(* IEC 61131-3 sources: IEC61131-3_ST_SCL_Mutation_Generator/Tests/mutatedCodeTraffic, 85 files *)

(* ---- M097.st ---- *)
FUNCTION_BLOCK TRAFFIC_CTRL

VAR_INPUT
    PedestrianButton1 : BOOL;
    PedestrianButton2 : BOOL;
END_VAR

VAR_OUTPUT
    NorthSouthRed : BOOL;
    NorthSouthYellow : BOOL;
    NorthSouthGreen : BOOL;
    EastWestRed : BOOL;
    EastWestYellow : BOOL;
    EastWestGreen : BOOL;
    PedestrianLight1 : BOOL;
    PedestrianLight2 : BOOL;
END_VAR

VAR
    LightState : INT := 0; (* 0: North-South Green, 1: North-South Yellow, 2: East-West Green, 3: East-West Yellow *)
    PedestrianRequest1 : BOOL := FALSE;
    PedestrianRequest2 : BOOL := FALSE;
    PedestrianCrossing : BOOL := FALSE;
    Timer : TON;
END_VAR

(* Check for pedestrian requests *)
IF PedestrianButton1 THEN
    PedestrianRequest1 := TRUE;
END_IF;

IF PedestrianButton2 THEN
    PedestrianRequest2 := TRUE;
END_IF;

(* Traffic light state machine *)
CASE LightState OF
    0: (* North-South Green *)
        NorthSouthGreen := TRUE;
        EastWestRed := TRUE;
        IF PedestrianRequest1 AND PedestrianRequest2 THEN (* MUTATED: LOGICAL_OP_REPLACE *)
            Timer(IN := TRUE, PT := T#2s); (* Pedestrian crossing grace period *)
            IF Timer.Q THEN
                Timer(IN := FALSE);
                LightState := 1;
            END_IF;
        END_IF;

    1: (* North-South Yellow *)
        NorthSouthYellow := TRUE;
        EastWestRed := TRUE;
        Timer(IN := TRUE, PT := T#2s); (* Yellow light duration *)
        IF Timer.Q THEN
            Timer(IN := FALSE);
            LightState := 2;
        END_IF;

    2: (* East-West Green *)
        EastWestGreen := TRUE;
        NorthSouthRed := TRUE;
        IF PedestrianRequest1 THEN
            PedestrianLight1 := TRUE;
            PedestrianCrossing := TRUE;
        END_IF;
        IF PedestrianRequest2 THEN
            PedestrianLight2 := TRUE;
            PedestrianCrossing := TRUE;
        END_IF;
        IF PedestrianCrossing THEN
            Timer(IN := TRUE, PT := T#2s); (* Pedestrian crossing period *)
            IF Timer.Q THEN
                Timer(IN := FALSE);
                PedestrianRequest1 := FALSE;
                PedestrianRequest2 := FALSE;
                PedestrianLight1 := FALSE;
                PedestrianLight2 := FALSE;
                PedestrianCrossing := FALSE;
                LightState := 3;
            END_IF;
        END_IF;

    3: (* East-West Yellow *)
        EastWestYellow := TRUE;
        NorthSouthRed := TRUE;
        Timer(IN := TRUE, PT := T#2s); (* Yellow light duration *)
        IF Timer.Q THEN
            Timer(IN := FALSE);
            LightState := 0;
        END_IF;

END_CASE;

END_FUNCTION_BLOCK

(* ---- M098.st ---- *)
FUNCTION_BLOCK TRAFFIC_CTRL

VAR_INPUT
    PedestrianButton1 : BOOL;
    PedestrianButton2 : BOOL;
END_VAR

VAR_OUTPUT
    NorthSouthRed : BOOL;
    NorthSouthYellow : BOOL;
    NorthSouthGreen : BOOL;
    EastWestRed : BOOL;
    EastWestYellow : BOOL;
    EastWestGreen : BOOL;
    PedestrianLight1 : BOOL;
    PedestrianLight2 : BOOL;
END_VAR

VAR
    LightState : INT := 0; (* 0: North-South Green, 1: North-South Yellow, 2: East-West Green, 3: East-West Yellow *)
    PedestrianRequest1 : BOOL := FALSE;
    PedestrianRequest2 : BOOL := FALSE;
    PedestrianCrossing : BOOL := FALSE;
    Timer : TON;
END_VAR

(* Check for pedestrian requests *)
IF PedestrianButton1 THEN
    PedestrianRequest1 := TRUE;
END_IF;

IF PedestrianButton2 THEN
    PedestrianRequest2 := TRUE;
END_IF;

(* Traffic light state machine *)
CASE LightState OF
    0: (* North+South Green *) (* MUTATED: ARITH_OP_REPLACE *)
        NorthSouthGreen := TRUE;
        EastWestRed := TRUE;
        IF PedestrianRequest1 OR PedestrianRequest2 THEN
            Timer(IN := TRUE, PT := T#2s); (* Pedestrian crossing grace period *)
            IF Timer.Q THEN
                Timer(IN := FALSE);
                LightState := 1;
            END_IF;
        END_IF;

    1: (* North-South Yellow *)
        NorthSouthYellow := TRUE;
        EastWestRed := TRUE;
        Timer(IN := TRUE, PT := T#2s); (* Yellow light duration *)
        IF Timer.Q THEN
            Timer(IN := FALSE);
            LightState := 2;
        END_IF;

    2: (* East-West Green *)
        EastWestGreen := TRUE;
        NorthSouthRed := TRUE;
        IF PedestrianRequest1 THEN
            PedestrianLight1 := TRUE;
            PedestrianCrossing := TRUE;
        END_IF;
        IF PedestrianRequest2 THEN
            PedestrianLight2 := TRUE;
            PedestrianCrossing := TRUE;
        END_IF;
        IF PedestrianCrossing THEN
            Timer(IN := TRUE, PT := T#2s); (* Pedestrian crossing period *)
            IF Timer.Q THEN
                Timer(IN := FALSE);
                PedestrianRequest1 := FALSE;
                PedestrianRequest2 := FALSE;
                PedestrianLight1 := FALSE;
                PedestrianLight2 := FALSE;
                PedestrianCrossing := FALSE;
                LightState := 3;
            END_IF;
        END_IF;

    3: (* East-West Yellow *)
        EastWestYellow := TRUE;
        NorthSouthRed := TRUE;
        Timer(IN := TRUE, PT := T#2s); (* Yellow light duration *)
        IF Timer.Q THEN
            Timer(IN := FALSE);
            LightState := 0;
        END_IF;

END_CASE;

END_FUNCTION_BLOCK

(* ---- M099.st ---- *)
FUNCTION_BLOCK TRAFFIC_CTRL

VAR_INPUT
    PedestrianButton1 : BOOL;
    PedestrianButton2 : BOOL;
END_VAR

VAR_OUTPUT
    NorthSouthRed : BOOL;
    NorthSouthYellow : BOOL;
    NorthSouthGreen : BOOL;
    EastWestRed : BOOL;
    EastWestYellow : BOOL;
    EastWestGreen : BOOL;
    PedestrianLight1 : BOOL;
    PedestrianLight2 : BOOL;
END_VAR

VAR
    LightState : INT := 0; (* 0: North-South Green, 1: North-South Yellow, 2: East-West Green, 3: East-West Yellow *)
    PedestrianRequest1 : BOOL := FALSE;
    PedestrianRequest2 : BOOL := FALSE;
    PedestrianCrossing : BOOL := FALSE;
    Timer : TON;
END_VAR

(* Check for pedestrian requests *)
IF PedestrianButton1 THEN
    PedestrianRequest1 := TRUE;
END_IF;

IF PedestrianButton2 THEN
    PedestrianRequest2 := TRUE;
END_IF;

(* Traffic light state machine *)
CASE LightState OF
    0: (* North-South Green *)
        NorthSouthGreen := TRUE;
        EastWestRed := TRUE;
        IF PedestrianRequest1 OR PedestrianRequest2 THEN
            Timer(IN := TRUE, PT := T#2s); (* Pedestrian crossing grace period *)
            IF Timer.Q THEN
                Timer(IN := FALSE);
                LightState := 1;
            END_IF;
        END_IF;

    1: (* North+South Yellow *) (* MUTATED: ARITH_OP_REPLACE *)
        NorthSouthYellow := TRUE;
        EastWestRed := TRUE;
        Timer(IN := TRUE, PT := T#2s); (* Yellow light duration *)
        IF Timer.Q THEN
            Timer(IN := FALSE);
            LightState := 2;
        END_IF;

    2: (* East-West Green *)
        EastWestGreen := TRUE;
        NorthSouthRed := TRUE;
        IF PedestrianRequest1 THEN
            PedestrianLight1 := TRUE;
            PedestrianCrossing := TRUE;
        END_IF;
        IF PedestrianRequest2 THEN
            PedestrianLight2 := TRUE;
            PedestrianCrossing := TRUE;
        END_IF;
        IF PedestrianCrossing THEN
            Timer(IN := TRUE, PT := T#2s); (* Pedestrian crossing period *)
            IF Timer.Q THEN
                Timer(IN := FALSE);
                PedestrianRequest1 := FALSE;
                PedestrianRequest2 := FALSE;
                PedestrianLight1 := FALSE;
                PedestrianLight2 := FALSE;
                PedestrianCrossing := FALSE;
                LightState := 3;
            END_IF;
        END_IF;

    3: (* East-West Yellow *)
        EastWestYellow := TRUE;
        NorthSouthRed := TRUE;
        Timer(IN := TRUE, PT := T#2s); (* Yellow light duration *)
        IF Timer.Q THEN
            Timer(IN := FALSE);
            LightState := 0;
        END_IF;

END_CASE;

END_FUNCTION_BLOCK

(* ---- M100.st ---- *)
FUNCTION_BLOCK TRAFFIC_CTRL

VAR_INPUT
    PedestrianButton1 : BOOL;
    PedestrianButton2 : BOOL;
END_VAR

VAR_OUTPUT
    NorthSouthRed : BOOL;
    NorthSouthYellow : BOOL;
    NorthSouthGreen : BOOL;
    EastWestRed : BOOL;
    EastWestYellow : BOOL;
    EastWestGreen : BOOL;
    PedestrianLight1 : BOOL;
    PedestrianLight2 : BOOL;
END_VAR

VAR
    LightState : INT := 0; (* 0: North-South Green, 1: North-South Yellow, 2: East-West Green, 3: East-West Yellow *)
    PedestrianRequest1 : BOOL := FALSE;
    PedestrianRequest2 : BOOL := FALSE;
    PedestrianCrossing : BOOL := FALSE;
    Timer : TON;
END_VAR

(* Check for pedestrian requests *)
IF PedestrianButton1 THEN
    PedestrianRequest1 := TRUE;
END_IF;

IF PedestrianButton2 THEN
    PedestrianRequest2 := TRUE;
END_IF;

(* Traffic light state machine *)
CASE LightState OF
    0: (* North-South Green *)
        NorthSouthGreen := TRUE;
        EastWestRed := TRUE;
        IF PedestrianRequest1 OR PedestrianRequest2 THEN
            Timer(IN := TRUE, PT := T#2s); (* Pedestrian crossing grace period *)
            IF Timer.Q THEN
                Timer(IN := FALSE);
                LightState := 1;
            END_IF;
        END_IF;

    1: (* North-South Yellow *)
        NorthSouthYellow := TRUE;
        EastWestRed := TRUE;
        Timer(IN := TRUE, PT := T#2s); (* Yellow light duration *)
        IF Timer.Q THEN
            Timer(IN := FALSE);
            LightState := 2;
        END_IF;

    2: (* East+West Green *) (* MUTATED: ARITH_OP_REPLACE *)
        EastWestGreen := TRUE;
        NorthSouthRed := TRUE;
        IF PedestrianRequest1 THEN
            PedestrianLight1 := TRUE;
            PedestrianCrossing := TRUE;
        END_IF;
        IF PedestrianRequest2 THEN
            PedestrianLight2 := TRUE;
            PedestrianCrossing := TRUE;
        END_IF;
        IF PedestrianCrossing THEN
            Timer(IN := TRUE, PT := T#2s); (* Pedestrian crossing period *)
            IF Timer.Q THEN
                Timer(IN := FALSE);
                PedestrianRequest1 := FALSE;
                PedestrianRequest2 := FALSE;
                PedestrianLight1 := FALSE;
                PedestrianLight2 := FALSE;
                PedestrianCrossing := FALSE;
                LightState := 3;
            END_IF;
        END_IF;

    3: (* East-West Yellow *)
        EastWestYellow := TRUE;
        NorthSouthRed := TRUE;
        Timer(IN := TRUE, PT := T#2s); (* Yellow light duration *)
        IF Timer.Q THEN
            Timer(IN := FALSE);
            LightState := 0;
        END_IF;

END_CASE;

END_FUNCTION_BLOCK

(* ---- M101.st ---- *)
FUNCTION_BLOCK TRAFFIC_CTRL

VAR_INPUT
    PedestrianButton1 : BOOL;
    PedestrianButton2 : BOOL;
END_VAR

VAR_OUTPUT
    NorthSouthRed : BOOL;
    NorthSouthYellow : BOOL;
    NorthSouthGreen : BOOL;
    EastWestRed : BOOL;
    EastWestYellow : BOOL;
    EastWestGreen : BOOL;
    PedestrianLight1 : BOOL;
    PedestrianLight2 : BOOL;
END_VAR

VAR
    LightState : INT := 0; (* 0: North-South Green, 1: North-South Yellow, 2: East-West Green, 3: East-West Yellow *)
    PedestrianRequest1 : BOOL := FALSE;
    PedestrianRequest2 : BOOL := FALSE;
    PedestrianCrossing : BOOL := FALSE;
    Timer : TON;
END_VAR

(* Check for pedestrian requests *)
IF PedestrianButton1 THEN
    PedestrianRequest1 := TRUE;
END_IF;

IF PedestrianButton2 THEN
    PedestrianRequest2 := TRUE;
END_IF;

(* Traffic light state machine *)
CASE LightState OF
    0: (* North-South Green *)
        NorthSouthGreen := TRUE;
        EastWestRed := TRUE;
        IF PedestrianRequest1 OR PedestrianRequest2 THEN
            Timer(IN := TRUE, PT := T#2s); (* Pedestrian crossing grace period *)
            IF Timer.Q THEN
                Timer(IN := FALSE);
                LightState := 1;
            END_IF;
        END_IF;

    1: (* North-South Yellow *)
        NorthSouthYellow := TRUE;
        EastWestRed := TRUE;
        Timer(IN := TRUE, PT := T#2s); (* Yellow light duration *)
        IF Timer.Q THEN
            Timer(IN := FALSE);
            LightState := 2;
        END_IF;

    2: (* East-West Green *)
        EastWestGreen := TRUE;
        NorthSouthRed := TRUE;
        IF PedestrianRequest1 THEN
            PedestrianLight1 := TRUE;
            PedestrianCrossing := TRUE;
        END_IF;
        IF PedestrianRequest2 THEN
            PedestrianLight2 := TRUE;
            PedestrianCrossing := TRUE;
        END_IF;
        IF PedestrianCrossing THEN
            Timer(IN := TRUE, PT := T#2s); (* Pedestrian crossing period *)
            IF Timer.Q THEN
                Timer(IN := FALSE);
                PedestrianRequest1 := FALSE;
                PedestrianRequest2 := FALSE;
                PedestrianLight1 := FALSE;
                PedestrianLight2 := FALSE;
                PedestrianCrossing := FALSE;
                LightState := 3;
            END_IF;
        END_IF;

    3: (* East+West Yellow *) (* MUTATED: ARITH_OP_REPLACE *)
        EastWestYellow := TRUE;
        NorthSouthRed := TRUE;
        Timer(IN := TRUE, PT := T#2s); (* Yellow light duration *)
        IF Timer.Q THEN
            Timer(IN := FALSE);
            LightState := 0;
        END_IF;

END_CASE;

END_FUNCTION_BLOCK

(* ---- M102.st ---- *)
FUNCTION_BLOCK TRAFFIC_CTRL

VAR_INPUT
    PedestrianButton1 : BOOL;
    PedestrianButton2 : BOOL;
END_VAR

VAR_OUTPUT
    NorthSouthRed : BOOL;
    NorthSouthYellow : BOOL;
    NorthSouthGreen : BOOL;
    EastWestRed : BOOL;
    EastWestYellow : BOOL;
    EastWestGreen : BOOL;
    PedestrianLight1 : BOOL;
    PedestrianLight2 : BOOL;
END_VAR

VAR
    LightState : INT := 0; (* 0: North-South Green, 1: North-South Yellow, 2: East-West Green, 3: East-West Yellow *)
    PedestrianRequest1 : BOOL := TRUE; (* MUTATED: BOOL_CONST_REPLACE *)
    PedestrianRequest2 : BOOL := FALSE;
    PedestrianCrossing : BOOL := FALSE;
    Timer : TON;
END_VAR

(* Check for pedestrian requests *)
IF PedestrianButton1 THEN
    PedestrianRequest1 := TRUE;
END_IF;

IF PedestrianButton2 THEN
    PedestrianRequest2 := TRUE;
END_IF;

(* Traffic light state machine *)
CASE LightState OF
    0: (* North-South Green *)
        NorthSouthGreen := TRUE;
        EastWestRed := TRUE;
        IF PedestrianRequest1 OR PedestrianRequest2 THEN
            Timer(IN := TRUE, PT := T#2s); (* Pedestrian crossing grace period *)
            IF Timer.Q THEN
                Timer(IN := FALSE);
                LightState := 1;
            END_IF;
        END_IF;

    1: (* North-South Yellow *)
        NorthSouthYellow := TRUE;
        EastWestRed := TRUE;
        Timer(IN := TRUE, PT := T#2s); (* Yellow light duration *)
        IF Timer.Q THEN
            Timer(IN := FALSE);
            LightState := 2;
        END_IF;

    2: (* East-West Green *)
        EastWestGreen := TRUE;
        NorthSouthRed := TRUE;
        IF PedestrianRequest1 THEN
            PedestrianLight1 := TRUE;
            PedestrianCrossing := TRUE;
        END_IF;
        IF PedestrianRequest2 THEN
            PedestrianLight2 := TRUE;
            PedestrianCrossing := TRUE;
        END_IF;
        IF PedestrianCrossing THEN
            Timer(IN := TRUE, PT := T#2s); (* Pedestrian crossing period *)
            IF Timer.Q THEN
                Timer(IN := FALSE);
                PedestrianRequest1 := FALSE;
                PedestrianRequest2 := FALSE;
                PedestrianLight1 := FALSE;
                PedestrianLight2 := FALSE;
                PedestrianCrossing := FALSE;
                LightState := 3;
            END_IF;
        END_IF;

    3: (* East-West Yellow *)
        EastWestYellow := TRUE;
        NorthSouthRed := TRUE;
        Timer(IN := TRUE, PT := T#2s); (* Yellow light duration *)
        IF Timer.Q THEN
            Timer(IN := FALSE);
            LightState := 0;
        END_IF;

END_CASE;

END_FUNCTION_BLOCK

(* ---- M103.st ---- *)
FUNCTION_BLOCK TRAFFIC_CTRL

VAR_INPUT
    PedestrianButton1 : BOOL;
    PedestrianButton2 : BOOL;
END_VAR

VAR_OUTPUT
    NorthSouthRed : BOOL;
    NorthSouthYellow : BOOL;
    NorthSouthGreen : BOOL;
    EastWestRed : BOOL;
    EastWestYellow : BOOL;
    EastWestGreen : BOOL;
    PedestrianLight1 : BOOL;
    PedestrianLight2 : BOOL;
END_VAR

VAR
    LightState : INT := 0; (* 0: North-South Green, 1: North-South Yellow, 2: East-West Green, 3: East-West Yellow *)
    PedestrianRequest1 : BOOL := FALSE;
    PedestrianRequest2 : BOOL := TRUE; (* MUTATED: BOOL_CONST_REPLACE *)
    PedestrianCrossing : BOOL := FALSE;
    Timer : TON;
END_VAR

(* Check for pedestrian requests *)
IF PedestrianButton1 THEN
    PedestrianRequest1 := TRUE;
END_IF;

IF PedestrianButton2 THEN
    PedestrianRequest2 := TRUE;
END_IF;

(* Traffic light state machine *)
CASE LightState OF
    0: (* North-South Green *)
        NorthSouthGreen := TRUE;
        EastWestRed := TRUE;
        IF PedestrianRequest1 OR PedestrianRequest2 THEN
            Timer(IN := TRUE, PT := T#2s); (* Pedestrian crossing grace period *)
            IF Timer.Q THEN
                Timer(IN := FALSE);
                LightState := 1;
            END_IF;
        END_IF;

    1: (* North-South Yellow *)
        NorthSouthYellow := TRUE;
        EastWestRed := TRUE;
        Timer(IN := TRUE, PT := T#2s); (* Yellow light duration *)
        IF Timer.Q THEN
            Timer(IN := FALSE);
            LightState := 2;
        END_IF;

    2: (* East-West Green *)
        EastWestGreen := TRUE;
        NorthSouthRed := TRUE;
        IF PedestrianRequest1 THEN
            PedestrianLight1 := TRUE;
            PedestrianCrossing := TRUE;
        END_IF;
        IF PedestrianRequest2 THEN
            PedestrianLight2 := TRUE;
            PedestrianCrossing := TRUE;
        END_IF;
        IF PedestrianCrossing THEN
            Timer(IN := TRUE, PT := T#2s); (* Pedestrian crossing period *)
            IF Timer.Q THEN
                Timer(IN := FALSE);
                PedestrianRequest1 := FALSE;
                PedestrianRequest2 := FALSE;
                PedestrianLight1 := FALSE;
                PedestrianLight2 := FALSE;
                PedestrianCrossing := FALSE;
                LightState := 3;
            END_IF;
        END_IF;

    3: (* East-West Yellow *)
        EastWestYellow := TRUE;
        NorthSouthRed := TRUE;
        Timer(IN := TRUE, PT := T#2s); (* Yellow light duration *)
        IF Timer.Q THEN
            Timer(IN := FALSE);
            LightState := 0;
        END_IF;

END_CASE;

END_FUNCTION_BLOCK

(* ---- M104.st ---- *)
FUNCTION_BLOCK TRAFFIC_CTRL

VAR_INPUT
    PedestrianButton1 : BOOL;
    PedestrianButton2 : BOOL;
END_VAR

VAR_OUTPUT
    NorthSouthRed : BOOL;
    NorthSouthYellow : BOOL;
    NorthSouthGreen : BOOL;
    EastWestRed : BOOL;
    EastWestYellow : BOOL;
    EastWestGreen : BOOL;
    PedestrianLight1 : BOOL;
    PedestrianLight2 : BOOL;
END_VAR

VAR
    LightState : INT := 0; (* 0: North-South Green, 1: North-South Yellow, 2: East-West Green, 3: East-West Yellow *)
    PedestrianRequest1 : BOOL := FALSE;
    PedestrianRequest2 : BOOL := FALSE;
    PedestrianCrossing : BOOL := TRUE; (* MUTATED: BOOL_CONST_REPLACE *)
    Timer : TON;
END_VAR

(* Check for pedestrian requests *)
IF PedestrianButton1 THEN
    PedestrianRequest1 := TRUE;
END_IF;

IF PedestrianButton2 THEN
    PedestrianRequest2 := TRUE;
END_IF;

(* Traffic light state machine *)
CASE LightState OF
    0: (* North-South Green *)
        NorthSouthGreen := TRUE;
        EastWestRed := TRUE;
        IF PedestrianRequest1 OR PedestrianRequest2 THEN
            Timer(IN := TRUE, PT := T#2s); (* Pedestrian crossing grace period *)
            IF Timer.Q THEN
                Timer(IN := FALSE);
                LightState := 1;
            END_IF;
        END_IF;

    1: (* North-South Yellow *)
        NorthSouthYellow := TRUE;
        EastWestRed := TRUE;
        Timer(IN := TRUE, PT := T#2s); (* Yellow light duration *)
        IF Timer.Q THEN
            Timer(IN := FALSE);
            LightState := 2;
        END_IF;

    2: (* East-West Green *)
        EastWestGreen := TRUE;
        NorthSouthRed := TRUE;
        IF PedestrianRequest1 THEN
            PedestrianLight1 := TRUE;
            PedestrianCrossing := TRUE;
        END_IF;
        IF PedestrianRequest2 THEN
            PedestrianLight2 := TRUE;
            PedestrianCrossing := TRUE;
        END_IF;
        IF PedestrianCrossing THEN
            Timer(IN := TRUE, PT := T#2s); (* Pedestrian crossing period *)
            IF Timer.Q THEN
                Timer(IN := FALSE);
                PedestrianRequest1 := FALSE;
                PedestrianRequest2 := FALSE;
                PedestrianLight1 := FALSE;
                PedestrianLight2 := FALSE;
                PedestrianCrossing := FALSE;
                LightState := 3;
            END_IF;
        END_IF;

    3: (* East-West Yellow *)
        EastWestYellow := TRUE;
        NorthSouthRed := TRUE;
        Timer(IN := TRUE, PT := T#2s); (* Yellow light duration *)
        IF Timer.Q THEN
            Timer(IN := FALSE);
            LightState := 0;
        END_IF;

END_CASE;

END_FUNCTION_BLOCK

(* ---- M105.st ---- *)
FUNCTION_BLOCK TRAFFIC_CTRL

VAR_INPUT
    PedestrianButton1 : BOOL;
    PedestrianButton2 : BOOL;
END_VAR

VAR_OUTPUT
    NorthSouthRed : BOOL;
    NorthSouthYellow : BOOL;
    NorthSouthGreen : BOOL;
    EastWestRed : BOOL;
    EastWestYellow : BOOL;
    EastWestGreen : BOOL;
    PedestrianLight1 : BOOL;
    PedestrianLight2 : BOOL;
END_VAR

VAR
    LightState : INT := 0; (* 0: North-South Green, 1: North-South Yellow, 2: East-West Green, 3: East-West Yellow *)
    PedestrianRequest1 : BOOL := FALSE;
    PedestrianRequest2 : BOOL := FALSE;
    PedestrianCrossing : BOOL := FALSE;
    Timer : TON;
END_VAR

(* Check for pedestrian requests *)
IF PedestrianButton1 THEN
    PedestrianRequest1 := FALSE; (* MUTATED: BOOL_CONST_REPLACE *)
END_IF;

IF PedestrianButton2 THEN
    PedestrianRequest2 := TRUE;
END_IF;

(* Traffic light state machine *)
CASE LightState OF
    0: (* North-South Green *)
        NorthSouthGreen := TRUE;
        EastWestRed := TRUE;
        IF PedestrianRequest1 OR PedestrianRequest2 THEN
            Timer(IN := TRUE, PT := T#2s); (* Pedestrian crossing grace period *)
            IF Timer.Q THEN
                Timer(IN := FALSE);
                LightState := 1;
            END_IF;
        END_IF;

    1: (* North-South Yellow *)
        NorthSouthYellow := TRUE;
        EastWestRed := TRUE;
        Timer(IN := TRUE, PT := T#2s); (* Yellow light duration *)
        IF Timer.Q THEN
            Timer(IN := FALSE);
            LightState := 2;
        END_IF;

    2: (* East-West Green *)
        EastWestGreen := TRUE;
        NorthSouthRed := TRUE;
        IF PedestrianRequest1 THEN
            PedestrianLight1 := TRUE;
            PedestrianCrossing := TRUE;
        END_IF;
        IF PedestrianRequest2 THEN
            PedestrianLight2 := TRUE;
            PedestrianCrossing := TRUE;
        END_IF;
        IF PedestrianCrossing THEN
            Timer(IN := TRUE, PT := T#2s); (* Pedestrian crossing period *)
            IF Timer.Q THEN
                Timer(IN := FALSE);
                PedestrianRequest1 := FALSE;
                PedestrianRequest2 := FALSE;
                PedestrianLight1 := FALSE;
                PedestrianLight2 := FALSE;
                PedestrianCrossing := FALSE;
                LightState := 3;
            END_IF;
        END_IF;

    3: (* East-West Yellow *)
        EastWestYellow := TRUE;
        NorthSouthRed := TRUE;
        Timer(IN := TRUE, PT := T#2s); (* Yellow light duration *)
        IF Timer.Q THEN
            Timer(IN := FALSE);
            LightState := 0;
        END_IF;

END_CASE;

END_FUNCTION_BLOCK

(* ---- M106.st ---- *)
FUNCTION_BLOCK TRAFFIC_CTRL

VAR_INPUT
    PedestrianButton1 : BOOL;
    PedestrianButton2 : BOOL;
END_VAR

VAR_OUTPUT
    NorthSouthRed : BOOL;
    NorthSouthYellow : BOOL;
    NorthSouthGreen : BOOL;
    EastWestRed : BOOL;
    EastWestYellow : BOOL;
    EastWestGreen : BOOL;
    PedestrianLight1 : BOOL;
    PedestrianLight2 : BOOL;
END_VAR

VAR
    LightState : INT := 0; (* 0: North-South Green, 1: North-South Yellow, 2: East-West Green, 3: East-West Yellow *)
    PedestrianRequest1 : BOOL := FALSE;
    PedestrianRequest2 : BOOL := FALSE;
    PedestrianCrossing : BOOL := FALSE;
    Timer : TON;
END_VAR

(* Check for pedestrian requests *)
IF PedestrianButton1 THEN
    PedestrianRequest1 := TRUE;
END_IF;

IF PedestrianButton2 THEN
    PedestrianRequest2 := FALSE; (* MUTATED: BOOL_CONST_REPLACE *)
END_IF;

(* Traffic light state machine *)
CASE LightState OF
    0: (* North-South Green *)
        NorthSouthGreen := TRUE;
        EastWestRed := TRUE;
        IF PedestrianRequest1 OR PedestrianRequest2 THEN
            Timer(IN := TRUE, PT := T#2s); (* Pedestrian crossing grace period *)
            IF Timer.Q THEN
                Timer(IN := FALSE);
                LightState := 1;
            END_IF;
        END_IF;

    1: (* North-South Yellow *)
        NorthSouthYellow := TRUE;
        EastWestRed := TRUE;
        Timer(IN := TRUE, PT := T#2s); (* Yellow light duration *)
        IF Timer.Q THEN
            Timer(IN := FALSE);
            LightState := 2;
        END_IF;

    2: (* East-West Green *)
        EastWestGreen := TRUE;
        NorthSouthRed := TRUE;
        IF PedestrianRequest1 THEN
            PedestrianLight1 := TRUE;
            PedestrianCrossing := TRUE;
        END_IF;
        IF PedestrianRequest2 THEN
            PedestrianLight2 := TRUE;
            PedestrianCrossing := TRUE;
        END_IF;
        IF PedestrianCrossing THEN
            Timer(IN := TRUE, PT := T#2s); (* Pedestrian crossing period *)
            IF Timer.Q THEN
                Timer(IN := FALSE);
                PedestrianRequest1 := FALSE;
                PedestrianRequest2 := FALSE;
                PedestrianLight1 := FALSE;
                PedestrianLight2 := FALSE;
                PedestrianCrossing := FALSE;
                LightState := 3;
            END_IF;
        END_IF;

    3: (* East-West Yellow *)
        EastWestYellow := TRUE;
        NorthSouthRed := TRUE;
        Timer(IN := TRUE, PT := T#2s); (* Yellow light duration *)
        IF Timer.Q THEN
            Timer(IN := FALSE);
            LightState := 0;
        END_IF;

END_CASE;

END_FUNCTION_BLOCK

(* ---- M107.st ---- *)
FUNCTION_BLOCK TRAFFIC_CTRL

VAR_INPUT
    PedestrianButton1 : BOOL;
    PedestrianButton2 : BOOL;
END_VAR

VAR_OUTPUT
    NorthSouthRed : BOOL;
    NorthSouthYellow : BOOL;
    NorthSouthGreen : BOOL;
    EastWestRed : BOOL;
    EastWestYellow : BOOL;
    EastWestGreen : BOOL;
    PedestrianLight1 : BOOL;
    PedestrianLight2 : BOOL;
END_VAR

VAR
    LightState : INT := 0; (* 0: North-South Green, 1: North-South Yellow, 2: East-West Green, 3: East-West Yellow *)
    PedestrianRequest1 : BOOL := FALSE;
    PedestrianRequest2 : BOOL := FALSE;
    PedestrianCrossing : BOOL := FALSE;
    Timer : TON;
END_VAR

(* Check for pedestrian requests *)
IF PedestrianButton1 THEN
    PedestrianRequest1 := TRUE;
END_IF;

IF PedestrianButton2 THEN
    PedestrianRequest2 := TRUE;
END_IF;

(* Traffic light state machine *)
CASE LightState OF
    0: (* North-South Green *)
        NorthSouthGreen := FALSE; (* MUTATED: BOOL_CONST_REPLACE *)
        EastWestRed := TRUE;
        IF PedestrianRequest1 OR PedestrianRequest2 THEN
            Timer(IN := TRUE, PT := T#2s); (* Pedestrian crossing grace period *)
            IF Timer.Q THEN
                Timer(IN := FALSE);
                LightState := 1;
            END_IF;
        END_IF;

    1: (* North-South Yellow *)
        NorthSouthYellow := TRUE;
        EastWestRed := TRUE;
        Timer(IN := TRUE, PT := T#2s); (* Yellow light duration *)
        IF Timer.Q THEN
            Timer(IN := FALSE);
            LightState := 2;
        END_IF;

    2: (* East-West Green *)
        EastWestGreen := TRUE;
        NorthSouthRed := TRUE;
        IF PedestrianRequest1 THEN
            PedestrianLight1 := TRUE;
            PedestrianCrossing := TRUE;
        END_IF;
        IF PedestrianRequest2 THEN
            PedestrianLight2 := TRUE;
            PedestrianCrossing := TRUE;
        END_IF;
        IF PedestrianCrossing THEN
            Timer(IN := TRUE, PT := T#2s); (* Pedestrian crossing period *)
            IF Timer.Q THEN
                Timer(IN := FALSE);
                PedestrianRequest1 := FALSE;
                PedestrianRequest2 := FALSE;
                PedestrianLight1 := FALSE;
                PedestrianLight2 := FALSE;
                PedestrianCrossing := FALSE;
                LightState := 3;
            END_IF;
        END_IF;

    3: (* East-West Yellow *)
        EastWestYellow := TRUE;
        NorthSouthRed := TRUE;
        Timer(IN := TRUE, PT := T#2s); (* Yellow light duration *)
        IF Timer.Q THEN
            Timer(IN := FALSE);
            LightState := 0;
        END_IF;

END_CASE;

END_FUNCTION_BLOCK

(* ---- M108.st ---- *)
FUNCTION_BLOCK TRAFFIC_CTRL

VAR_INPUT
    PedestrianButton1 : BOOL;
    PedestrianButton2 : BOOL;
END_VAR

VAR_OUTPUT
    NorthSouthRed : BOOL;
    NorthSouthYellow : BOOL;
    NorthSouthGreen : BOOL;
    EastWestRed : BOOL;
    EastWestYellow : BOOL;
    EastWestGreen : BOOL;
    PedestrianLight1 : BOOL;
    PedestrianLight2 : BOOL;
END_VAR

VAR
    LightState : INT := 0; (* 0: North-South Green, 1: North-South Yellow, 2: East-West Green, 3: East-West Yellow *)
    PedestrianRequest1 : BOOL := FALSE;
    PedestrianRequest2 : BOOL := FALSE;
    PedestrianCrossing : BOOL := FALSE;
    Timer : TON;
END_VAR

(* Check for pedestrian requests *)
IF PedestrianButton1 THEN
    PedestrianRequest1 := TRUE;
END_IF;

IF PedestrianButton2 THEN
    PedestrianRequest2 := TRUE;
END_IF;

(* Traffic light state machine *)
CASE LightState OF
    0: (* North-South Green *)
        NorthSouthGreen := TRUE;
        EastWestRed := FALSE; (* MUTATED: BOOL_CONST_REPLACE *)
        IF PedestrianRequest1 OR PedestrianRequest2 THEN
            Timer(IN := TRUE, PT := T#2s); (* Pedestrian crossing grace period *)
            IF Timer.Q THEN
                Timer(IN := FALSE);
                LightState := 1;
            END_IF;
        END_IF;

    1: (* North-South Yellow *)
        NorthSouthYellow := TRUE;
        EastWestRed := TRUE;
        Timer(IN := TRUE, PT := T#2s); (* Yellow light duration *)
        IF Timer.Q THEN
            Timer(IN := FALSE);
            LightState := 2;
        END_IF;

    2: (* East-West Green *)
        EastWestGreen := TRUE;
        NorthSouthRed := TRUE;
        IF PedestrianRequest1 THEN
            PedestrianLight1 := TRUE;
            PedestrianCrossing := TRUE;
        END_IF;
        IF PedestrianRequest2 THEN
            PedestrianLight2 := TRUE;
            PedestrianCrossing := TRUE;
        END_IF;
        IF PedestrianCrossing THEN
            Timer(IN := TRUE, PT := T#2s); (* Pedestrian crossing period *)
            IF Timer.Q THEN
                Timer(IN := FALSE);
                PedestrianRequest1 := FALSE;
                PedestrianRequest2 := FALSE;
                PedestrianLight1 := FALSE;
                PedestrianLight2 := FALSE;
                PedestrianCrossing := FALSE;
                LightState := 3;
            END_IF;
        END_IF;

    3: (* East-West Yellow *)
        EastWestYellow := TRUE;
        NorthSouthRed := TRUE;
        Timer(IN := TRUE, PT := T#2s); (* Yellow light duration *)
        IF Timer.Q THEN
            Timer(IN := FALSE);
            LightState := 0;
        END_IF;

END_CASE;

END_FUNCTION_BLOCK

(* ---- M109.st ---- *)
FUNCTION_BLOCK TRAFFIC_CTRL

VAR_INPUT
    PedestrianButton1 : BOOL;
    PedestrianButton2 : BOOL;
END_VAR

VAR_OUTPUT
    NorthSouthRed : BOOL;
    NorthSouthYellow : BOOL;
    NorthSouthGreen : BOOL;
    EastWestRed : BOOL;
    EastWestYellow : BOOL;
    EastWestGreen : BOOL;
    PedestrianLight1 : BOOL;
    PedestrianLight2 : BOOL;
END_VAR

VAR
    LightState : INT := 0; (* 0: North-South Green, 1: North-South Yellow, 2: East-West Green, 3: East-West Yellow *)
    PedestrianRequest1 : BOOL := FALSE;
    PedestrianRequest2 : BOOL := FALSE;
    PedestrianCrossing : BOOL := FALSE;
    Timer : TON;
END_VAR

(* Check for pedestrian requests *)
IF PedestrianButton1 THEN
    PedestrianRequest1 := TRUE;
END_IF;

IF PedestrianButton2 THEN
    PedestrianRequest2 := TRUE;
END_IF;

(* Traffic light state machine *)
CASE LightState OF
    0: (* North-South Green *)
        NorthSouthGreen := TRUE;
        EastWestRed := TRUE;
        IF PedestrianRequest1 OR PedestrianRequest2 THEN
            Timer(IN := FALSE, PT := T#2s); (* Pedestrian crossing grace period *) (* MUTATED: BOOL_CONST_REPLACE *)
            IF Timer.Q THEN
                Timer(IN := FALSE);
                LightState := 1;
            END_IF;
        END_IF;

    1: (* North-South Yellow *)
        NorthSouthYellow := TRUE;
        EastWestRed := TRUE;
        Timer(IN := TRUE, PT := T#2s); (* Yellow light duration *)
        IF Timer.Q THEN
            Timer(IN := FALSE);
            LightState := 2;
        END_IF;

    2: (* East-West Green *)
        EastWestGreen := TRUE;
        NorthSouthRed := TRUE;
        IF PedestrianRequest1 THEN
            PedestrianLight1 := TRUE;
            PedestrianCrossing := TRUE;
        END_IF;
        IF PedestrianRequest2 THEN
            PedestrianLight2 := TRUE;
            PedestrianCrossing := TRUE;
        END_IF;
        IF PedestrianCrossing THEN
            Timer(IN := TRUE, PT := T#2s); (* Pedestrian crossing period *)
            IF Timer.Q THEN
                Timer(IN := FALSE);
                PedestrianRequest1 := FALSE;
                PedestrianRequest2 := FALSE;
                PedestrianLight1 := FALSE;
                PedestrianLight2 := FALSE;
                PedestrianCrossing := FALSE;
                LightState := 3;
            END_IF;
        END_IF;

    3: (* East-West Yellow *)
        EastWestYellow := TRUE;
        NorthSouthRed := TRUE;
        Timer(IN := TRUE, PT := T#2s); (* Yellow light duration *)
        IF Timer.Q THEN
            Timer(IN := FALSE);
            LightState := 0;
        END_IF;

END_CASE;

END_FUNCTION_BLOCK

(* ---- M110.st ---- *)
FUNCTION_BLOCK TRAFFIC_CTRL

VAR_INPUT
    PedestrianButton1 : BOOL;
    PedestrianButton2 : BOOL;
END_VAR

VAR_OUTPUT
    NorthSouthRed : BOOL;
    NorthSouthYellow : BOOL;
    NorthSouthGreen : BOOL;
    EastWestRed : BOOL;
    EastWestYellow : BOOL;
    EastWestGreen : BOOL;
    PedestrianLight1 : BOOL;
    PedestrianLight2 : BOOL;
END_VAR

VAR
    LightState : INT := 0; (* 0: North-South Green, 1: North-South Yellow, 2: East-West Green, 3: East-West Yellow *)
    PedestrianRequest1 : BOOL := FALSE;
    PedestrianRequest2 : BOOL := FALSE;
    PedestrianCrossing : BOOL := FALSE;
    Timer : TON;
END_VAR

(* Check for pedestrian requests *)
IF PedestrianButton1 THEN
    PedestrianRequest1 := TRUE;
END_IF;

IF PedestrianButton2 THEN
    PedestrianRequest2 := TRUE;
END_IF;

(* Traffic light state machine *)
CASE LightState OF
    0: (* North-South Green *)
        NorthSouthGreen := TRUE;
        EastWestRed := TRUE;
        IF PedestrianRequest1 OR PedestrianRequest2 THEN
            Timer(IN := TRUE, PT := T#2s); (* Pedestrian crossing grace period *)
            IF Timer.Q THEN
                Timer(IN := TRUE); (* MUTATED: BOOL_CONST_REPLACE *)
                LightState := 1;
            END_IF;
        END_IF;

    1: (* North-South Yellow *)
        NorthSouthYellow := TRUE;
        EastWestRed := TRUE;
        Timer(IN := TRUE, PT := T#2s); (* Yellow light duration *)
        IF Timer.Q THEN
            Timer(IN := FALSE);
            LightState := 2;
        END_IF;

    2: (* East-West Green *)
        EastWestGreen := TRUE;
        NorthSouthRed := TRUE;
        IF PedestrianRequest1 THEN
            PedestrianLight1 := TRUE;
            PedestrianCrossing := TRUE;
        END_IF;
        IF PedestrianRequest2 THEN
            PedestrianLight2 := TRUE;
            PedestrianCrossing := TRUE;
        END_IF;
        IF PedestrianCrossing THEN
            Timer(IN := TRUE, PT := T#2s); (* Pedestrian crossing period *)
            IF Timer.Q THEN
                Timer(IN := FALSE);
                PedestrianRequest1 := FALSE;
                PedestrianRequest2 := FALSE;
                PedestrianLight1 := FALSE;
                PedestrianLight2 := FALSE;
                PedestrianCrossing := FALSE;
                LightState := 3;
            END_IF;
        END_IF;

    3: (* East-West Yellow *)
        EastWestYellow := TRUE;
        NorthSouthRed := TRUE;
        Timer(IN := TRUE, PT := T#2s); (* Yellow light duration *)
        IF Timer.Q THEN
            Timer(IN := FALSE);
            LightState := 0;
        END_IF;

END_CASE;

END_FUNCTION_BLOCK

(* ---- M111.st ---- *)
FUNCTION_BLOCK TRAFFIC_CTRL

VAR_INPUT
    PedestrianButton1 : BOOL;
    PedestrianButton2 : BOOL;
END_VAR

VAR_OUTPUT
    NorthSouthRed : BOOL;
    NorthSouthYellow : BOOL;
    NorthSouthGreen : BOOL;
    EastWestRed : BOOL;
    EastWestYellow : BOOL;
    EastWestGreen : BOOL;
    PedestrianLight1 : BOOL;
    PedestrianLight2 : BOOL;
END_VAR

VAR
    LightState : INT := 0; (* 0: North-South Green, 1: North-South Yellow, 2: East-West Green, 3: East-West Yellow *)
    PedestrianRequest1 : BOOL := FALSE;
    PedestrianRequest2 : BOOL := FALSE;
    PedestrianCrossing : BOOL := FALSE;
    Timer : TON;
END_VAR

(* Check for pedestrian requests *)
IF PedestrianButton1 THEN
    PedestrianRequest1 := TRUE;
END_IF;

IF PedestrianButton2 THEN
    PedestrianRequest2 := TRUE;
END_IF;

(* Traffic light state machine *)
CASE LightState OF
    0: (* North-South Green *)
        NorthSouthGreen := TRUE;
        EastWestRed := TRUE;
        IF PedestrianRequest1 OR PedestrianRequest2 THEN
            Timer(IN := TRUE, PT := T#2s); (* Pedestrian crossing grace period *)
            IF Timer.Q THEN
                Timer(IN := FALSE);
                LightState := 1;
            END_IF;
        END_IF;

    1: (* North-South Yellow *)
        NorthSouthYellow := FALSE; (* MUTATED: BOOL_CONST_REPLACE *)
        EastWestRed := TRUE;
        Timer(IN := TRUE, PT := T#2s); (* Yellow light duration *)
        IF Timer.Q THEN
            Timer(IN := FALSE);
            LightState := 2;
        END_IF;

    2: (* East-West Green *)
        EastWestGreen := TRUE;
        NorthSouthRed := TRUE;
        IF PedestrianRequest1 THEN
            PedestrianLight1 := TRUE;
            PedestrianCrossing := TRUE;
        END_IF;
        IF PedestrianRequest2 THEN
            PedestrianLight2 := TRUE;
            PedestrianCrossing := TRUE;
        END_IF;
        IF PedestrianCrossing THEN
            Timer(IN := TRUE, PT := T#2s); (* Pedestrian crossing period *)
            IF Timer.Q THEN
                Timer(IN := FALSE);
                PedestrianRequest1 := FALSE;
                PedestrianRequest2 := FALSE;
                PedestrianLight1 := FALSE;
                PedestrianLight2 := FALSE;
                PedestrianCrossing := FALSE;
                LightState := 3;
            END_IF;
        END_IF;

    3: (* East-West Yellow *)
        EastWestYellow := TRUE;
        NorthSouthRed := TRUE;
        Timer(IN := TRUE, PT := T#2s); (* Yellow light duration *)
        IF Timer.Q THEN
            Timer(IN := FALSE);
            LightState := 0;
        END_IF;

END_CASE;

END_FUNCTION_BLOCK

(* ---- M112.st ---- *)
FUNCTION_BLOCK TRAFFIC_CTRL

VAR_INPUT
    PedestrianButton1 : BOOL;
    PedestrianButton2 : BOOL;
END_VAR

VAR_OUTPUT
    NorthSouthRed : BOOL;
    NorthSouthYellow : BOOL;
    NorthSouthGreen : BOOL;
    EastWestRed : BOOL;
    EastWestYellow : BOOL;
    EastWestGreen : BOOL;
    PedestrianLight1 : BOOL;
    PedestrianLight2 : BOOL;
END_VAR

VAR
    LightState : INT := 0; (* 0: North-South Green, 1: North-South Yellow, 2: East-West Green, 3: East-West Yellow *)
    PedestrianRequest1 : BOOL := FALSE;
    PedestrianRequest2 : BOOL := FALSE;
    PedestrianCrossing : BOOL := FALSE;
    Timer : TON;
END_VAR

(* Check for pedestrian requests *)
IF PedestrianButton1 THEN
    PedestrianRequest1 := TRUE;
END_IF;

IF PedestrianButton2 THEN
    PedestrianRequest2 := TRUE;
END_IF;

(* Traffic light state machine *)
CASE LightState OF
    0: (* North-South Green *)
        NorthSouthGreen := TRUE;
        EastWestRed := TRUE;
        IF PedestrianRequest1 OR PedestrianRequest2 THEN
            Timer(IN := TRUE, PT := T#2s); (* Pedestrian crossing grace period *)
            IF Timer.Q THEN
                Timer(IN := FALSE);
                LightState := 1;
            END_IF;
        END_IF;

    1: (* North-South Yellow *)
        NorthSouthYellow := TRUE;
        EastWestRed := FALSE; (* MUTATED: BOOL_CONST_REPLACE *)
        Timer(IN := TRUE, PT := T#2s); (* Yellow light duration *)
        IF Timer.Q THEN
            Timer(IN := FALSE);
            LightState := 2;
        END_IF;

    2: (* East-West Green *)
        EastWestGreen := TRUE;
        NorthSouthRed := TRUE;
        IF PedestrianRequest1 THEN
            PedestrianLight1 := TRUE;
            PedestrianCrossing := TRUE;
        END_IF;
        IF PedestrianRequest2 THEN
            PedestrianLight2 := TRUE;
            PedestrianCrossing := TRUE;
        END_IF;
        IF PedestrianCrossing THEN
            Timer(IN := TRUE, PT := T#2s); (* Pedestrian crossing period *)
            IF Timer.Q THEN
                Timer(IN := FALSE);
                PedestrianRequest1 := FALSE;
                PedestrianRequest2 := FALSE;
                PedestrianLight1 := FALSE;
                PedestrianLight2 := FALSE;
                PedestrianCrossing := FALSE;
                LightState := 3;
            END_IF;
        END_IF;

    3: (* East-West Yellow *)
        EastWestYellow := TRUE;
        NorthSouthRed := TRUE;
        Timer(IN := TRUE, PT := T#2s); (* Yellow light duration *)
        IF Timer.Q THEN
            Timer(IN := FALSE);
            LightState := 0;
        END_IF;

END_CASE;

END_FUNCTION_BLOCK

(* ---- M113.st ---- *)
FUNCTION_BLOCK TRAFFIC_CTRL

VAR_INPUT
    PedestrianButton1 : BOOL;
    PedestrianButton2 : BOOL;
END_VAR

VAR_OUTPUT
    NorthSouthRed : BOOL;
    NorthSouthYellow : BOOL;
    NorthSouthGreen : BOOL;
    EastWestRed : BOOL;
    EastWestYellow : BOOL;
    EastWestGreen : BOOL;
    PedestrianLight1 : BOOL;
    PedestrianLight2 : BOOL;
END_VAR

VAR
    LightState : INT := 0; (* 0: North-South Green, 1: North-South Yellow, 2: East-West Green, 3: East-West Yellow *)
    PedestrianRequest1 : BOOL := FALSE;
    PedestrianRequest2 : BOOL := FALSE;
    PedestrianCrossing : BOOL := FALSE;
    Timer : TON;
END_VAR

(* Check for pedestrian requests *)
IF PedestrianButton1 THEN
    PedestrianRequest1 := TRUE;
END_IF;

IF PedestrianButton2 THEN
    PedestrianRequest2 := TRUE;
END_IF;

(* Traffic light state machine *)
CASE LightState OF
    0: (* North-South Green *)
        NorthSouthGreen := TRUE;
        EastWestRed := TRUE;
        IF PedestrianRequest1 OR PedestrianRequest2 THEN
            Timer(IN := TRUE, PT := T#2s); (* Pedestrian crossing grace period *)
            IF Timer.Q THEN
                Timer(IN := FALSE);
                LightState := 1;
            END_IF;
        END_IF;

    1: (* North-South Yellow *)
        NorthSouthYellow := TRUE;
        EastWestRed := TRUE;
        Timer(IN := FALSE, PT := T#2s); (* Yellow light duration *) (* MUTATED: BOOL_CONST_REPLACE *)
        IF Timer.Q THEN
            Timer(IN := FALSE);
            LightState := 2;
        END_IF;

    2: (* East-West Green *)
        EastWestGreen := TRUE;
        NorthSouthRed := TRUE;
        IF PedestrianRequest1 THEN
            PedestrianLight1 := TRUE;
            PedestrianCrossing := TRUE;
        END_IF;
        IF PedestrianRequest2 THEN
            PedestrianLight2 := TRUE;
            PedestrianCrossing := TRUE;
        END_IF;
        IF PedestrianCrossing THEN
            Timer(IN := TRUE, PT := T#2s); (* Pedestrian crossing period *)
            IF Timer.Q THEN
                Timer(IN := FALSE);
                PedestrianRequest1 := FALSE;
                PedestrianRequest2 := FALSE;
                PedestrianLight1 := FALSE;
                PedestrianLight2 := FALSE;
                PedestrianCrossing := FALSE;
                LightState := 3;
            END_IF;
        END_IF;

    3: (* East-West Yellow *)
        EastWestYellow := TRUE;
        NorthSouthRed := TRUE;
        Timer(IN := TRUE, PT := T#2s); (* Yellow light duration *)
        IF Timer.Q THEN
            Timer(IN := FALSE);
            LightState := 0;
        END_IF;

END_CASE;

END_FUNCTION_BLOCK

(* ---- M114.st ---- *)
FUNCTION_BLOCK TRAFFIC_CTRL

VAR_INPUT
    PedestrianButton1 : BOOL;
    PedestrianButton2 : BOOL;
END_VAR

VAR_OUTPUT
    NorthSouthRed : BOOL;
    NorthSouthYellow : BOOL;
    NorthSouthGreen : BOOL;
    EastWestRed : BOOL;
    EastWestYellow : BOOL;
    EastWestGreen : BOOL;
    PedestrianLight1 : BOOL;
    PedestrianLight2 : BOOL;
END_VAR

VAR
    LightState : INT := 0; (* 0: North-South Green, 1: North-South Yellow, 2: East-West Green, 3: East-West Yellow *)
    PedestrianRequest1 : BOOL := FALSE;
    PedestrianRequest2 : BOOL := FALSE;
    PedestrianCrossing : BOOL := FALSE;
    Timer : TON;
END_VAR

(* Check for pedestrian requests *)
IF PedestrianButton1 THEN
    PedestrianRequest1 := TRUE;
END_IF;

IF PedestrianButton2 THEN
    PedestrianRequest2 := TRUE;
END_IF;

(* Traffic light state machine *)
CASE LightState OF
    0: (* North-South Green *)
        NorthSouthGreen := TRUE;
        EastWestRed := TRUE;
        IF PedestrianRequest1 OR PedestrianRequest2 THEN
            Timer(IN := TRUE, PT := T#2s); (* Pedestrian crossing grace period *)
            IF Timer.Q THEN
                Timer(IN := FALSE);
                LightState := 1;
            END_IF;
        END_IF;

    1: (* North-South Yellow *)
        NorthSouthYellow := TRUE;
        EastWestRed := TRUE;
        Timer(IN := TRUE, PT := T#2s); (* Yellow light duration *)
        IF Timer.Q THEN
            Timer(IN := TRUE); (* MUTATED: BOOL_CONST_REPLACE *)
            LightState := 2;
        END_IF;

    2: (* East-West Green *)
        EastWestGreen := TRUE;
        NorthSouthRed := TRUE;
        IF PedestrianRequest1 THEN
            PedestrianLight1 := TRUE;
            PedestrianCrossing := TRUE;
        END_IF;
        IF PedestrianRequest2 THEN
            PedestrianLight2 := TRUE;
            PedestrianCrossing := TRUE;
        END_IF;
        IF PedestrianCrossing THEN
            Timer(IN := TRUE, PT := T#2s); (* Pedestrian crossing period *)
            IF Timer.Q THEN
                Timer(IN := FALSE);
                PedestrianRequest1 := FALSE;
                PedestrianRequest2 := FALSE;
                PedestrianLight1 := FALSE;
                PedestrianLight2 := FALSE;
                PedestrianCrossing := FALSE;
                LightState := 3;
            END_IF;
        END_IF;

    3: (* East-West Yellow *)
        EastWestYellow := TRUE;
        NorthSouthRed := TRUE;
        Timer(IN := TRUE, PT := T#2s); (* Yellow light duration *)
        IF Timer.Q THEN
            Timer(IN := FALSE);
            LightState := 0;
        END_IF;

END_CASE;

END_FUNCTION_BLOCK

(* ---- M115.st ---- *)
FUNCTION_BLOCK TRAFFIC_CTRL

VAR_INPUT
    PedestrianButton1 : BOOL;
    PedestrianButton2 : BOOL;
END_VAR

VAR_OUTPUT
    NorthSouthRed : BOOL;
    NorthSouthYellow : BOOL;
    NorthSouthGreen : BOOL;
    EastWestRed : BOOL;
    EastWestYellow : BOOL;
    EastWestGreen : BOOL;
    PedestrianLight1 : BOOL;
    PedestrianLight2 : BOOL;
END_VAR

VAR
    LightState : INT := 0; (* 0: North-South Green, 1: North-South Yellow, 2: East-West Green, 3: East-West Yellow *)
    PedestrianRequest1 : BOOL := FALSE;
    PedestrianRequest2 : BOOL := FALSE;
    PedestrianCrossing : BOOL := FALSE;
    Timer : TON;
END_VAR

(* Check for pedestrian requests *)
IF PedestrianButton1 THEN
    PedestrianRequest1 := TRUE;
END_IF;

IF PedestrianButton2 THEN
    PedestrianRequest2 := TRUE;
END_IF;

(* Traffic light state machine *)
CASE LightState OF
    0: (* North-South Green *)
        NorthSouthGreen := TRUE;
        EastWestRed := TRUE;
        IF PedestrianRequest1 OR PedestrianRequest2 THEN
            Timer(IN := TRUE, PT := T#2s); (* Pedestrian crossing grace period *)
            IF Timer.Q THEN
                Timer(IN := FALSE);
                LightState := 1;
            END_IF;
        END_IF;

    1: (* North-South Yellow *)
        NorthSouthYellow := TRUE;
        EastWestRed := TRUE;
        Timer(IN := TRUE, PT := T#2s); (* Yellow light duration *)
        IF Timer.Q THEN
            Timer(IN := FALSE);
            LightState := 2;
        END_IF;

    2: (* East-West Green *)
        EastWestGreen := FALSE; (* MUTATED: BOOL_CONST_REPLACE *)
        NorthSouthRed := TRUE;
        IF PedestrianRequest1 THEN
            PedestrianLight1 := TRUE;
            PedestrianCrossing := TRUE;
        END_IF;
        IF PedestrianRequest2 THEN
            PedestrianLight2 := TRUE;
            PedestrianCrossing := TRUE;
        END_IF;
        IF PedestrianCrossing THEN
            Timer(IN := TRUE, PT := T#2s); (* Pedestrian crossing period *)
            IF Timer.Q THEN
                Timer(IN := FALSE);
                PedestrianRequest1 := FALSE;
                PedestrianRequest2 := FALSE;
                PedestrianLight1 := FALSE;
                PedestrianLight2 := FALSE;
                PedestrianCrossing := FALSE;
                LightState := 3;
            END_IF;
        END_IF;

    3: (* East-West Yellow *)
        EastWestYellow := TRUE;
        NorthSouthRed := TRUE;
        Timer(IN := TRUE, PT := T#2s); (* Yellow light duration *)
        IF Timer.Q THEN
            Timer(IN := FALSE);
            LightState := 0;
        END_IF;

END_CASE;

END_FUNCTION_BLOCK

(* ---- M116.st ---- *)
FUNCTION_BLOCK TRAFFIC_CTRL

VAR_INPUT
    PedestrianButton1 : BOOL;
    PedestrianButton2 : BOOL;
END_VAR

VAR_OUTPUT
    NorthSouthRed : BOOL;
    NorthSouthYellow : BOOL;
    NorthSouthGreen : BOOL;
    EastWestRed : BOOL;
    EastWestYellow : BOOL;
    EastWestGreen : BOOL;
    PedestrianLight1 : BOOL;
    PedestrianLight2 : BOOL;
END_VAR

VAR
    LightState : INT := 0; (* 0: North-South Green, 1: North-South Yellow, 2: East-West Green, 3: East-West Yellow *)
    PedestrianRequest1 : BOOL := FALSE;
    PedestrianRequest2 : BOOL := FALSE;
    PedestrianCrossing : BOOL := FALSE;
    Timer : TON;
END_VAR

(* Check for pedestrian requests *)
IF PedestrianButton1 THEN
    PedestrianRequest1 := TRUE;
END_IF;

IF PedestrianButton2 THEN
    PedestrianRequest2 := TRUE;
END_IF;

(* Traffic light state machine *)
CASE LightState OF
    0: (* North-South Green *)
        NorthSouthGreen := TRUE;
        EastWestRed := TRUE;
        IF PedestrianRequest1 OR PedestrianRequest2 THEN
            Timer(IN := TRUE, PT := T#2s); (* Pedestrian crossing grace period *)
            IF Timer.Q THEN
                Timer(IN := FALSE);
                LightState := 1;
            END_IF;
        END_IF;

    1: (* North-South Yellow *)
        NorthSouthYellow := TRUE;
        EastWestRed := TRUE;
        Timer(IN := TRUE, PT := T#2s); (* Yellow light duration *)
        IF Timer.Q THEN
            Timer(IN := FALSE);
            LightState := 2;
        END_IF;

    2: (* East-West Green *)
        EastWestGreen := TRUE;
        NorthSouthRed := FALSE; (* MUTATED: BOOL_CONST_REPLACE *)
        IF PedestrianRequest1 THEN
            PedestrianLight1 := TRUE;
            PedestrianCrossing := TRUE;
        END_IF;
        IF PedestrianRequest2 THEN
            PedestrianLight2 := TRUE;
            PedestrianCrossing := TRUE;
        END_IF;
        IF PedestrianCrossing THEN
            Timer(IN := TRUE, PT := T#2s); (* Pedestrian crossing period *)
            IF Timer.Q THEN
                Timer(IN := FALSE);
                PedestrianRequest1 := FALSE;
                PedestrianRequest2 := FALSE;
                PedestrianLight1 := FALSE;
                PedestrianLight2 := FALSE;
                PedestrianCrossing := FALSE;
                LightState := 3;
            END_IF;
        END_IF;

    3: (* East-West Yellow *)
        EastWestYellow := TRUE;
        NorthSouthRed := TRUE;
        Timer(IN := TRUE, PT := T#2s); (* Yellow light duration *)
        IF Timer.Q THEN
            Timer(IN := FALSE);
            LightState := 0;
        END_IF;

END_CASE;

END_FUNCTION_BLOCK

(* ---- M117.st ---- *)
FUNCTION_BLOCK TRAFFIC_CTRL

VAR_INPUT
    PedestrianButton1 : BOOL;
    PedestrianButton2 : BOOL;
END_VAR

VAR_OUTPUT
    NorthSouthRed : BOOL;
    NorthSouthYellow : BOOL;
    NorthSouthGreen : BOOL;
    EastWestRed : BOOL;
    EastWestYellow : BOOL;
    EastWestGreen : BOOL;
    PedestrianLight1 : BOOL;
    PedestrianLight2 : BOOL;
END_VAR

VAR
    LightState : INT := 0; (* 0: North-South Green, 1: North-South Yellow, 2: East-West Green, 3: East-West Yellow *)
    PedestrianRequest1 : BOOL := FALSE;
    PedestrianRequest2 : BOOL := FALSE;
    PedestrianCrossing : BOOL := FALSE;
    Timer : TON;
END_VAR

(* Check for pedestrian requests *)
IF PedestrianButton1 THEN
    PedestrianRequest1 := TRUE;
END_IF;

IF PedestrianButton2 THEN
    PedestrianRequest2 := TRUE;
END_IF;

(* Traffic light state machine *)
CASE LightState OF
    0: (* North-South Green *)
        NorthSouthGreen := TRUE;
        EastWestRed := TRUE;
        IF PedestrianRequest1 OR PedestrianRequest2 THEN
            Timer(IN := TRUE, PT := T#2s); (* Pedestrian crossing grace period *)
            IF Timer.Q THEN
                Timer(IN := FALSE);
                LightState := 1;
            END_IF;
        END_IF;

    1: (* North-South Yellow *)
        NorthSouthYellow := TRUE;
        EastWestRed := TRUE;
        Timer(IN := TRUE, PT := T#2s); (* Yellow light duration *)
        IF Timer.Q THEN
            Timer(IN := FALSE);
            LightState := 2;
        END_IF;

    2: (* East-West Green *)
        EastWestGreen := TRUE;
        NorthSouthRed := TRUE;
        IF PedestrianRequest1 THEN
            PedestrianLight1 := FALSE; (* MUTATED: BOOL_CONST_REPLACE *)
            PedestrianCrossing := TRUE;
        END_IF;
        IF PedestrianRequest2 THEN
            PedestrianLight2 := TRUE;
            PedestrianCrossing := TRUE;
        END_IF;
        IF PedestrianCrossing THEN
            Timer(IN := TRUE, PT := T#2s); (* Pedestrian crossing period *)
            IF Timer.Q THEN
                Timer(IN := FALSE);
                PedestrianRequest1 := FALSE;
                PedestrianRequest2 := FALSE;
                PedestrianLight1 := FALSE;
                PedestrianLight2 := FALSE;
                PedestrianCrossing := FALSE;
                LightState := 3;
            END_IF;
        END_IF;

    3: (* East-West Yellow *)
        EastWestYellow := TRUE;
        NorthSouthRed := TRUE;
        Timer(IN := TRUE, PT := T#2s); (* Yellow light duration *)
        IF Timer.Q THEN
            Timer(IN := FALSE);
            LightState := 0;
        END_IF;

END_CASE;

END_FUNCTION_BLOCK

(* ---- M118.st ---- *)
FUNCTION_BLOCK TRAFFIC_CTRL

VAR_INPUT
    PedestrianButton1 : BOOL;
    PedestrianButton2 : BOOL;
END_VAR

VAR_OUTPUT
    NorthSouthRed : BOOL;
    NorthSouthYellow : BOOL;
    NorthSouthGreen : BOOL;
    EastWestRed : BOOL;
    EastWestYellow : BOOL;
    EastWestGreen : BOOL;
    PedestrianLight1 : BOOL;
    PedestrianLight2 : BOOL;
END_VAR

VAR
    LightState : INT := 0; (* 0: North-South Green, 1: North-South Yellow, 2: East-West Green, 3: East-West Yellow *)
    PedestrianRequest1 : BOOL := FALSE;
    PedestrianRequest2 : BOOL := FALSE;
    PedestrianCrossing : BOOL := FALSE;
    Timer : TON;
END_VAR

(* Check for pedestrian requests *)
IF PedestrianButton1 THEN
    PedestrianRequest1 := TRUE;
END_IF;

IF PedestrianButton2 THEN
    PedestrianRequest2 := TRUE;
END_IF;

(* Traffic light state machine *)
CASE LightState OF
    0: (* North-South Green *)
        NorthSouthGreen := TRUE;
        EastWestRed := TRUE;
        IF PedestrianRequest1 OR PedestrianRequest2 THEN
            Timer(IN := TRUE, PT := T#2s); (* Pedestrian crossing grace period *)
            IF Timer.Q THEN
                Timer(IN := FALSE);
                LightState := 1;
            END_IF;
        END_IF;

    1: (* North-South Yellow *)
        NorthSouthYellow := TRUE;
        EastWestRed := TRUE;
        Timer(IN := TRUE, PT := T#2s); (* Yellow light duration *)
        IF Timer.Q THEN
            Timer(IN := FALSE);
            LightState := 2;
        END_IF;

    2: (* East-West Green *)
        EastWestGreen := TRUE;
        NorthSouthRed := TRUE;
        IF PedestrianRequest1 THEN
            PedestrianLight1 := TRUE;
            PedestrianCrossing := FALSE; (* MUTATED: BOOL_CONST_REPLACE *)
        END_IF;
        IF PedestrianRequest2 THEN
            PedestrianLight2 := TRUE;
            PedestrianCrossing := TRUE;
        END_IF;
        IF PedestrianCrossing THEN
            Timer(IN := TRUE, PT := T#2s); (* Pedestrian crossing period *)
            IF Timer.Q THEN
                Timer(IN := FALSE);
                PedestrianRequest1 := FALSE;
                PedestrianRequest2 := FALSE;
                PedestrianLight1 := FALSE;
                PedestrianLight2 := FALSE;
                PedestrianCrossing := FALSE;
                LightState := 3;
            END_IF;
        END_IF;

    3: (* East-West Yellow *)
        EastWestYellow := TRUE;
        NorthSouthRed := TRUE;
        Timer(IN := TRUE, PT := T#2s); (* Yellow light duration *)
        IF Timer.Q THEN
            Timer(IN := FALSE);
            LightState := 0;
        END_IF;

END_CASE;

END_FUNCTION_BLOCK

(* ---- M119.st ---- *)
FUNCTION_BLOCK TRAFFIC_CTRL

VAR_INPUT
    PedestrianButton1 : BOOL;
    PedestrianButton2 : BOOL;
END_VAR

VAR_OUTPUT
    NorthSouthRed : BOOL;
    NorthSouthYellow : BOOL;
    NorthSouthGreen : BOOL;
    EastWestRed : BOOL;
    EastWestYellow : BOOL;
    EastWestGreen : BOOL;
    PedestrianLight1 : BOOL;
    PedestrianLight2 : BOOL;
END_VAR

VAR
    LightState : INT := 0; (* 0: North-South Green, 1: North-South Yellow, 2: East-West Green, 3: East-West Yellow *)
    PedestrianRequest1 : BOOL := FALSE;
    PedestrianRequest2 : BOOL := FALSE;
    PedestrianCrossing : BOOL := FALSE;
    Timer : TON;
END_VAR

(* Check for pedestrian requests *)
IF PedestrianButton1 THEN
    PedestrianRequest1 := TRUE;
END_IF;

IF PedestrianButton2 THEN
    PedestrianRequest2 := TRUE;
END_IF;

(* Traffic light state machine *)
CASE LightState OF
    0: (* North-South Green *)
        NorthSouthGreen := TRUE;
        EastWestRed := TRUE;
        IF PedestrianRequest1 OR PedestrianRequest2 THEN
            Timer(IN := TRUE, PT := T#2s); (* Pedestrian crossing grace period *)
            IF Timer.Q THEN
                Timer(IN := FALSE);
                LightState := 1;
            END_IF;
        END_IF;

    1: (* North-South Yellow *)
        NorthSouthYellow := TRUE;
        EastWestRed := TRUE;
        Timer(IN := TRUE, PT := T#2s); (* Yellow light duration *)
        IF Timer.Q THEN
            Timer(IN := FALSE);
            LightState := 2;
        END_IF;

    2: (* East-West Green *)
        EastWestGreen := TRUE;
        NorthSouthRed := TRUE;
        IF PedestrianRequest1 THEN
            PedestrianLight1 := TRUE;
            PedestrianCrossing := TRUE;
        END_IF;
        IF PedestrianRequest2 THEN
            PedestrianLight2 := FALSE; (* MUTATED: BOOL_CONST_REPLACE *)
            PedestrianCrossing := TRUE;
        END_IF;
        IF PedestrianCrossing THEN
            Timer(IN := TRUE, PT := T#2s); (* Pedestrian crossing period *)
            IF Timer.Q THEN
                Timer(IN := FALSE);
                PedestrianRequest1 := FALSE;
                PedestrianRequest2 := FALSE;
                PedestrianLight1 := FALSE;
                PedestrianLight2 := FALSE;
                PedestrianCrossing := FALSE;
                LightState := 3;
            END_IF;
        END_IF;

    3: (* East-West Yellow *)
        EastWestYellow := TRUE;
        NorthSouthRed := TRUE;
        Timer(IN := TRUE, PT := T#2s); (* Yellow light duration *)
        IF Timer.Q THEN
            Timer(IN := FALSE);
            LightState := 0;
        END_IF;

END_CASE;

END_FUNCTION_BLOCK

(* ---- M120.st ---- *)
FUNCTION_BLOCK TRAFFIC_CTRL

VAR_INPUT
    PedestrianButton1 : BOOL;
    PedestrianButton2 : BOOL;
END_VAR

VAR_OUTPUT
    NorthSouthRed : BOOL;
    NorthSouthYellow : BOOL;
    NorthSouthGreen : BOOL;
    EastWestRed : BOOL;
    EastWestYellow : BOOL;
    EastWestGreen : BOOL;
    PedestrianLight1 : BOOL;
    PedestrianLight2 : BOOL;
END_VAR

VAR
    LightState : INT := 0; (* 0: North-South Green, 1: North-South Yellow, 2: East-West Green, 3: East-West Yellow *)
    PedestrianRequest1 : BOOL := FALSE;
    PedestrianRequest2 : BOOL := FALSE;
    PedestrianCrossing : BOOL := FALSE;
    Timer : TON;
END_VAR

(* Check for pedestrian requests *)
IF PedestrianButton1 THEN
    PedestrianRequest1 := TRUE;
END_IF;

IF PedestrianButton2 THEN
    PedestrianRequest2 := TRUE;
END_IF;

(* Traffic light state machine *)
CASE LightState OF
    0: (* North-South Green *)
        NorthSouthGreen := TRUE;
        EastWestRed := TRUE;
        IF PedestrianRequest1 OR PedestrianRequest2 THEN
            Timer(IN := TRUE, PT := T#2s); (* Pedestrian crossing grace period *)
            IF Timer.Q THEN
                Timer(IN := FALSE);
                LightState := 1;
            END_IF;
        END_IF;

    1: (* North-South Yellow *)
        NorthSouthYellow := TRUE;
        EastWestRed := TRUE;
        Timer(IN := TRUE, PT := T#2s); (* Yellow light duration *)
        IF Timer.Q THEN
            Timer(IN := FALSE);
            LightState := 2;
        END_IF;

    2: (* East-West Green *)
        EastWestGreen := TRUE;
        NorthSouthRed := TRUE;
        IF PedestrianRequest1 THEN
            PedestrianLight1 := TRUE;
            PedestrianCrossing := TRUE;
        END_IF;
        IF PedestrianRequest2 THEN
            PedestrianLight2 := TRUE;
            PedestrianCrossing := FALSE; (* MUTATED: BOOL_CONST_REPLACE *)
        END_IF;
        IF PedestrianCrossing THEN
            Timer(IN := TRUE, PT := T#2s); (* Pedestrian crossing period *)
            IF Timer.Q THEN
                Timer(IN := FALSE);
                PedestrianRequest1 := FALSE;
                PedestrianRequest2 := FALSE;
                PedestrianLight1 := FALSE;
                PedestrianLight2 := FALSE;
                PedestrianCrossing := FALSE;
                LightState := 3;
            END_IF;
        END_IF;

    3: (* East-West Yellow *)
        EastWestYellow := TRUE;
        NorthSouthRed := TRUE;
        Timer(IN := TRUE, PT := T#2s); (* Yellow light duration *)
        IF Timer.Q THEN
            Timer(IN := FALSE);
            LightState := 0;
        END_IF;

END_CASE;

END_FUNCTION_BLOCK

(* ---- M121.st ---- *)
FUNCTION_BLOCK TRAFFIC_CTRL

VAR_INPUT
    PedestrianButton1 : BOOL;
    PedestrianButton2 : BOOL;
END_VAR

VAR_OUTPUT
    NorthSouthRed : BOOL;
    NorthSouthYellow : BOOL;
    NorthSouthGreen : BOOL;
    EastWestRed : BOOL;
    EastWestYellow : BOOL;
    EastWestGreen : BOOL;
    PedestrianLight1 : BOOL;
    PedestrianLight2 : BOOL;
END_VAR

VAR
    LightState : INT := 0; (* 0: North-South Green, 1: North-South Yellow, 2: East-West Green, 3: East-West Yellow *)
    PedestrianRequest1 : BOOL := FALSE;
    PedestrianRequest2 : BOOL := FALSE;
    PedestrianCrossing : BOOL := FALSE;
    Timer : TON;
END_VAR

(* Check for pedestrian requests *)
IF PedestrianButton1 THEN
    PedestrianRequest1 := TRUE;
END_IF;

IF PedestrianButton2 THEN
    PedestrianRequest2 := TRUE;
END_IF;

(* Traffic light state machine *)
CASE LightState OF
    0: (* North-South Green *)
        NorthSouthGreen := TRUE;
        EastWestRed := TRUE;
        IF PedestrianRequest1 OR PedestrianRequest2 THEN
            Timer(IN := TRUE, PT := T#2s); (* Pedestrian crossing grace period *)
            IF Timer.Q THEN
                Timer(IN := FALSE);
                LightState := 1;
            END_IF;
        END_IF;

    1: (* North-South Yellow *)
        NorthSouthYellow := TRUE;
        EastWestRed := TRUE;
        Timer(IN := TRUE, PT := T#2s); (* Yellow light duration *)
        IF Timer.Q THEN
            Timer(IN := FALSE);
            LightState := 2;
        END_IF;

    2: (* East-West Green *)
        EastWestGreen := TRUE;
        NorthSouthRed := TRUE;
        IF PedestrianRequest1 THEN
            PedestrianLight1 := TRUE;
            PedestrianCrossing := TRUE;
        END_IF;
        IF PedestrianRequest2 THEN
            PedestrianLight2 := TRUE;
            PedestrianCrossing := TRUE;
        END_IF;
        IF PedestrianCrossing THEN
            Timer(IN := FALSE, PT := T#2s); (* Pedestrian crossing period *) (* MUTATED: BOOL_CONST_REPLACE *)
            IF Timer.Q THEN
                Timer(IN := FALSE);
                PedestrianRequest1 := FALSE;
                PedestrianRequest2 := FALSE;
                PedestrianLight1 := FALSE;
                PedestrianLight2 := FALSE;
                PedestrianCrossing := FALSE;
                LightState := 3;
            END_IF;
        END_IF;

    3: (* East-West Yellow *)
        EastWestYellow := TRUE;
        NorthSouthRed := TRUE;
        Timer(IN := TRUE, PT := T#2s); (* Yellow light duration *)
        IF Timer.Q THEN
            Timer(IN := FALSE);
            LightState := 0;
        END_IF;

END_CASE;

END_FUNCTION_BLOCK

(* ---- M122.st ---- *)
FUNCTION_BLOCK TRAFFIC_CTRL

VAR_INPUT
    PedestrianButton1 : BOOL;
    PedestrianButton2 : BOOL;
END_VAR

VAR_OUTPUT
    NorthSouthRed : BOOL;
    NorthSouthYellow : BOOL;
    NorthSouthGreen : BOOL;
    EastWestRed : BOOL;
    EastWestYellow : BOOL;
    EastWestGreen : BOOL;
    PedestrianLight1 : BOOL;
    PedestrianLight2 : BOOL;
END_VAR

VAR
    LightState : INT := 0; (* 0: North-South Green, 1: North-South Yellow, 2: East-West Green, 3: East-West Yellow *)
    PedestrianRequest1 : BOOL := FALSE;
    PedestrianRequest2 : BOOL := FALSE;
    PedestrianCrossing : BOOL := FALSE;
    Timer : TON;
END_VAR

(* Check for pedestrian requests *)
IF PedestrianButton1 THEN
    PedestrianRequest1 := TRUE;
END_IF;

IF PedestrianButton2 THEN
    PedestrianRequest2 := TRUE;
END_IF;

(* Traffic light state machine *)
CASE LightState OF
    0: (* North-South Green *)
        NorthSouthGreen := TRUE;
        EastWestRed := TRUE;
        IF PedestrianRequest1 OR PedestrianRequest2 THEN
            Timer(IN := TRUE, PT := T#2s); (* Pedestrian crossing grace period *)
            IF Timer.Q THEN
                Timer(IN := FALSE);
                LightState := 1;
            END_IF;
        END_IF;

    1: (* North-South Yellow *)
        NorthSouthYellow := TRUE;
        EastWestRed := TRUE;
        Timer(IN := TRUE, PT := T#2s); (* Yellow light duration *)
        IF Timer.Q THEN
            Timer(IN := FALSE);
            LightState := 2;
        END_IF;

    2: (* East-West Green *)
        EastWestGreen := TRUE;
        NorthSouthRed := TRUE;
        IF PedestrianRequest1 THEN
            PedestrianLight1 := TRUE;
            PedestrianCrossing := TRUE;
        END_IF;
        IF PedestrianRequest2 THEN
            PedestrianLight2 := TRUE;
            PedestrianCrossing := TRUE;
        END_IF;
        IF PedestrianCrossing THEN
            Timer(IN := TRUE, PT := T#2s); (* Pedestrian crossing period *)
            IF Timer.Q THEN
                Timer(IN := TRUE); (* MUTATED: BOOL_CONST_REPLACE *)
                PedestrianRequest1 := FALSE;
                PedestrianRequest2 := FALSE;
                PedestrianLight1 := FALSE;
                PedestrianLight2 := FALSE;
                PedestrianCrossing := FALSE;
                LightState := 3;
            END_IF;
        END_IF;

    3: (* East-West Yellow *)
        EastWestYellow := TRUE;
        NorthSouthRed := TRUE;
        Timer(IN := TRUE, PT := T#2s); (* Yellow light duration *)
        IF Timer.Q THEN
            Timer(IN := FALSE);
            LightState := 0;
        END_IF;

END_CASE;

END_FUNCTION_BLOCK

(* ---- M123.st ---- *)
FUNCTION_BLOCK TRAFFIC_CTRL

VAR_INPUT
    PedestrianButton1 : BOOL;
    PedestrianButton2 : BOOL;
END_VAR

VAR_OUTPUT
    NorthSouthRed : BOOL;
    NorthSouthYellow : BOOL;
    NorthSouthGreen : BOOL;
    EastWestRed : BOOL;
    EastWestYellow : BOOL;
    EastWestGreen : BOOL;
    PedestrianLight1 : BOOL;
    PedestrianLight2 : BOOL;
END_VAR

VAR
    LightState : INT := 0; (* 0: North-South Green, 1: North-South Yellow, 2: East-West Green, 3: East-West Yellow *)
    PedestrianRequest1 : BOOL := FALSE;
    PedestrianRequest2 : BOOL := FALSE;
    PedestrianCrossing : BOOL := FALSE;
    Timer : TON;
END_VAR

(* Check for pedestrian requests *)
IF PedestrianButton1 THEN
    PedestrianRequest1 := TRUE;
END_IF;

IF PedestrianButton2 THEN
    PedestrianRequest2 := TRUE;
END_IF;

(* Traffic light state machine *)
CASE LightState OF
    0: (* North-South Green *)
        NorthSouthGreen := TRUE;
        EastWestRed := TRUE;
        IF PedestrianRequest1 OR PedestrianRequest2 THEN
            Timer(IN := TRUE, PT := T#2s); (* Pedestrian crossing grace period *)
            IF Timer.Q THEN
                Timer(IN := FALSE);
                LightState := 1;
            END_IF;
        END_IF;

    1: (* North-South Yellow *)
        NorthSouthYellow := TRUE;
        EastWestRed := TRUE;
        Timer(IN := TRUE, PT := T#2s); (* Yellow light duration *)
        IF Timer.Q THEN
            Timer(IN := FALSE);
            LightState := 2;
        END_IF;

    2: (* East-West Green *)
        EastWestGreen := TRUE;
        NorthSouthRed := TRUE;
        IF PedestrianRequest1 THEN
            PedestrianLight1 := TRUE;
            PedestrianCrossing := TRUE;
        END_IF;
        IF PedestrianRequest2 THEN
            PedestrianLight2 := TRUE;
            PedestrianCrossing := TRUE;
        END_IF;
        IF PedestrianCrossing THEN
            Timer(IN := TRUE, PT := T#2s); (* Pedestrian crossing period *)
            IF Timer.Q THEN
                Timer(IN := FALSE);
                PedestrianRequest1 := TRUE; (* MUTATED: BOOL_CONST_REPLACE *)
                PedestrianRequest2 := FALSE;
                PedestrianLight1 := FALSE;
                PedestrianLight2 := FALSE;
                PedestrianCrossing := FALSE;
                LightState := 3;
            END_IF;
        END_IF;

    3: (* East-West Yellow *)
        EastWestYellow := TRUE;
        NorthSouthRed := TRUE;
        Timer(IN := TRUE, PT := T#2s); (* Yellow light duration *)
        IF Timer.Q THEN
            Timer(IN := FALSE);
            LightState := 0;
        END_IF;

END_CASE;

END_FUNCTION_BLOCK

(* ---- M124.st ---- *)
FUNCTION_BLOCK TRAFFIC_CTRL

VAR_INPUT
    PedestrianButton1 : BOOL;
    PedestrianButton2 : BOOL;
END_VAR

VAR_OUTPUT
    NorthSouthRed : BOOL;
    NorthSouthYellow : BOOL;
    NorthSouthGreen : BOOL;
    EastWestRed : BOOL;
    EastWestYellow : BOOL;
    EastWestGreen : BOOL;
    PedestrianLight1 : BOOL;
    PedestrianLight2 : BOOL;
END_VAR

VAR
    LightState : INT := 0; (* 0: North-South Green, 1: North-South Yellow, 2: East-West Green, 3: East-West Yellow *)
    PedestrianRequest1 : BOOL := FALSE;
    PedestrianRequest2 : BOOL := FALSE;
    PedestrianCrossing : BOOL := FALSE;
    Timer : TON;
END_VAR

(* Check for pedestrian requests *)
IF PedestrianButton1 THEN
    PedestrianRequest1 := TRUE;
END_IF;

IF PedestrianButton2 THEN
    PedestrianRequest2 := TRUE;
END_IF;

(* Traffic light state machine *)
CASE LightState OF
    0: (* North-South Green *)
        NorthSouthGreen := TRUE;
        EastWestRed := TRUE;
        IF PedestrianRequest1 OR PedestrianRequest2 THEN
            Timer(IN := TRUE, PT := T#2s); (* Pedestrian crossing grace period *)
            IF Timer.Q THEN
                Timer(IN := FALSE);
                LightState := 1;
            END_IF;
        END_IF;

    1: (* North-South Yellow *)
        NorthSouthYellow := TRUE;
        EastWestRed := TRUE;
        Timer(IN := TRUE, PT := T#2s); (* Yellow light duration *)
        IF Timer.Q THEN
            Timer(IN := FALSE);
            LightState := 2;
        END_IF;

    2: (* East-West Green *)
        EastWestGreen := TRUE;
        NorthSouthRed := TRUE;
        IF PedestrianRequest1 THEN
            PedestrianLight1 := TRUE;
            PedestrianCrossing := TRUE;
        END_IF;
        IF PedestrianRequest2 THEN
            PedestrianLight2 := TRUE;
            PedestrianCrossing := TRUE;
        END_IF;
        IF PedestrianCrossing THEN
            Timer(IN := TRUE, PT := T#2s); (* Pedestrian crossing period *)
            IF Timer.Q THEN
                Timer(IN := FALSE);
                PedestrianRequest1 := FALSE;
                PedestrianRequest2 := TRUE; (* MUTATED: BOOL_CONST_REPLACE *)
                PedestrianLight1 := FALSE;
                PedestrianLight2 := FALSE;
                PedestrianCrossing := FALSE;
                LightState := 3;
            END_IF;
        END_IF;

    3: (* East-West Yellow *)
        EastWestYellow := TRUE;
        NorthSouthRed := TRUE;
        Timer(IN := TRUE, PT := T#2s); (* Yellow light duration *)
        IF Timer.Q THEN
            Timer(IN := FALSE);
            LightState := 0;
        END_IF;

END_CASE;

END_FUNCTION_BLOCK

(* ---- M125.st ---- *)
FUNCTION_BLOCK TRAFFIC_CTRL

VAR_INPUT
    PedestrianButton1 : BOOL;
    PedestrianButton2 : BOOL;
END_VAR

VAR_OUTPUT
    NorthSouthRed : BOOL;
    NorthSouthYellow : BOOL;
    NorthSouthGreen : BOOL;
    EastWestRed : BOOL;
    EastWestYellow : BOOL;
    EastWestGreen : BOOL;
    PedestrianLight1 : BOOL;
    PedestrianLight2 : BOOL;
END_VAR

VAR
    LightState : INT := 0; (* 0: North-South Green, 1: North-South Yellow, 2: East-West Green, 3: East-West Yellow *)
    PedestrianRequest1 : BOOL := FALSE;
    PedestrianRequest2 : BOOL := FALSE;
    PedestrianCrossing : BOOL := FALSE;
    Timer : TON;
END_VAR

(* Check for pedestrian requests *)
IF PedestrianButton1 THEN
    PedestrianRequest1 := TRUE;
END_IF;

IF PedestrianButton2 THEN
    PedestrianRequest2 := TRUE;
END_IF;

(* Traffic light state machine *)
CASE LightState OF
    0: (* North-South Green *)
        NorthSouthGreen := TRUE;
        EastWestRed := TRUE;
        IF PedestrianRequest1 OR PedestrianRequest2 THEN
            Timer(IN := TRUE, PT := T#2s); (* Pedestrian crossing grace period *)
            IF Timer.Q THEN
                Timer(IN := FALSE);
                LightState := 1;
            END_IF;
        END_IF;

    1: (* North-South Yellow *)
        NorthSouthYellow := TRUE;
        EastWestRed := TRUE;
        Timer(IN := TRUE, PT := T#2s); (* Yellow light duration *)
        IF Timer.Q THEN
            Timer(IN := FALSE);
            LightState := 2;
        END_IF;

    2: (* East-West Green *)
        EastWestGreen := TRUE;
        NorthSouthRed := TRUE;
        IF PedestrianRequest1 THEN
            PedestrianLight1 := TRUE;
            PedestrianCrossing := TRUE;
        END_IF;
        IF PedestrianRequest2 THEN
            PedestrianLight2 := TRUE;
            PedestrianCrossing := TRUE;
        END_IF;
        IF PedestrianCrossing THEN
            Timer(IN := TRUE, PT := T#2s); (* Pedestrian crossing period *)
            IF Timer.Q THEN
                Timer(IN := FALSE);
                PedestrianRequest1 := FALSE;
                PedestrianRequest2 := FALSE;
                PedestrianLight1 := TRUE; (* MUTATED: BOOL_CONST_REPLACE *)
                PedestrianLight2 := FALSE;
                PedestrianCrossing := FALSE;
                LightState := 3;
            END_IF;
        END_IF;

    3: (* East-West Yellow *)
        EastWestYellow := TRUE;
        NorthSouthRed := TRUE;
        Timer(IN := TRUE, PT := T#2s); (* Yellow light duration *)
        IF Timer.Q THEN
            Timer(IN := FALSE);
            LightState := 0;
        END_IF;

END_CASE;

END_FUNCTION_BLOCK

(* ---- M126.st ---- *)
FUNCTION_BLOCK TRAFFIC_CTRL

VAR_INPUT
    PedestrianButton1 : BOOL;
    PedestrianButton2 : BOOL;
END_VAR

VAR_OUTPUT
    NorthSouthRed : BOOL;
    NorthSouthYellow : BOOL;
    NorthSouthGreen : BOOL;
    EastWestRed : BOOL;
    EastWestYellow : BOOL;
    EastWestGreen : BOOL;
    PedestrianLight1 : BOOL;
    PedestrianLight2 : BOOL;
END_VAR

VAR
    LightState : INT := 0; (* 0: North-South Green, 1: North-South Yellow, 2: East-West Green, 3: East-West Yellow *)
    PedestrianRequest1 : BOOL := FALSE;
    PedestrianRequest2 : BOOL := FALSE;
    PedestrianCrossing : BOOL := FALSE;
    Timer : TON;
END_VAR

(* Check for pedestrian requests *)
IF PedestrianButton1 THEN
    PedestrianRequest1 := TRUE;
END_IF;

IF PedestrianButton2 THEN
    PedestrianRequest2 := TRUE;
END_IF;

(* Traffic light state machine *)
CASE LightState OF
    0: (* North-South Green *)
        NorthSouthGreen := TRUE;
        EastWestRed := TRUE;
        IF PedestrianRequest1 OR PedestrianRequest2 THEN
            Timer(IN := TRUE, PT := T#2s); (* Pedestrian crossing grace period *)
            IF Timer.Q THEN
                Timer(IN := FALSE);
                LightState := 1;
            END_IF;
        END_IF;

    1: (* North-South Yellow *)
        NorthSouthYellow := TRUE;
        EastWestRed := TRUE;
        Timer(IN := TRUE, PT := T#2s); (* Yellow light duration *)
        IF Timer.Q THEN
            Timer(IN := FALSE);
            LightState := 2;
        END_IF;

    2: (* East-West Green *)
        EastWestGreen := TRUE;
        NorthSouthRed := TRUE;
        IF PedestrianRequest1 THEN
            PedestrianLight1 := TRUE;
            PedestrianCrossing := TRUE;
        END_IF;
        IF PedestrianRequest2 THEN
            PedestrianLight2 := TRUE;
            PedestrianCrossing := TRUE;
        END_IF;
        IF PedestrianCrossing THEN
            Timer(IN := TRUE, PT := T#2s); (* Pedestrian crossing period *)
            IF Timer.Q THEN
                Timer(IN := FALSE);
                PedestrianRequest1 := FALSE;
                PedestrianRequest2 := FALSE;
                PedestrianLight1 := FALSE;
                PedestrianLight2 := TRUE; (* MUTATED: BOOL_CONST_REPLACE *)
                PedestrianCrossing := FALSE;
                LightState := 3;
            END_IF;
        END_IF;

    3: (* East-West Yellow *)
        EastWestYellow := TRUE;
        NorthSouthRed := TRUE;
        Timer(IN := TRUE, PT := T#2s); (* Yellow light duration *)
        IF Timer.Q THEN
            Timer(IN := FALSE);
            LightState := 0;
        END_IF;

END_CASE;

END_FUNCTION_BLOCK

(* ---- M127.st ---- *)
FUNCTION_BLOCK TRAFFIC_CTRL

VAR_INPUT
    PedestrianButton1 : BOOL;
    PedestrianButton2 : BOOL;
END_VAR

VAR_OUTPUT
    NorthSouthRed : BOOL;
    NorthSouthYellow : BOOL;
    NorthSouthGreen : BOOL;
    EastWestRed : BOOL;
    EastWestYellow : BOOL;
    EastWestGreen : BOOL;
    PedestrianLight1 : BOOL;
    PedestrianLight2 : BOOL;
END_VAR

VAR
    LightState : INT := 0; (* 0: North-South Green, 1: North-South Yellow, 2: East-West Green, 3: East-West Yellow *)
    PedestrianRequest1 : BOOL := FALSE;
    PedestrianRequest2 : BOOL := FALSE;
    PedestrianCrossing : BOOL := FALSE;
    Timer : TON;
END_VAR

(* Check for pedestrian requests *)
IF PedestrianButton1 THEN
    PedestrianRequest1 := TRUE;
END_IF;

IF PedestrianButton2 THEN
    PedestrianRequest2 := TRUE;
END_IF;

(* Traffic light state machine *)
CASE LightState OF
    0: (* North-South Green *)
        NorthSouthGreen := TRUE;
        EastWestRed := TRUE;
        IF PedestrianRequest1 OR PedestrianRequest2 THEN
            Timer(IN := TRUE, PT := T#2s); (* Pedestrian crossing grace period *)
            IF Timer.Q THEN
                Timer(IN := FALSE);
                LightState := 1;
            END_IF;
        END_IF;

    1: (* North-South Yellow *)
        NorthSouthYellow := TRUE;
        EastWestRed := TRUE;
        Timer(IN := TRUE, PT := T#2s); (* Yellow light duration *)
        IF Timer.Q THEN
            Timer(IN := FALSE);
            LightState := 2;
        END_IF;

    2: (* East-West Green *)
        EastWestGreen := TRUE;
        NorthSouthRed := TRUE;
        IF PedestrianRequest1 THEN
            PedestrianLight1 := TRUE;
            PedestrianCrossing := TRUE;
        END_IF;
        IF PedestrianRequest2 THEN
            PedestrianLight2 := TRUE;
            PedestrianCrossing := TRUE;
        END_IF;
        IF PedestrianCrossing THEN
            Timer(IN := TRUE, PT := T#2s); (* Pedestrian crossing period *)
            IF Timer.Q THEN
                Timer(IN := FALSE);
                PedestrianRequest1 := FALSE;
                PedestrianRequest2 := FALSE;
                PedestrianLight1 := FALSE;
                PedestrianLight2 := FALSE;
                PedestrianCrossing := TRUE; (* MUTATED: BOOL_CONST_REPLACE *)
                LightState := 3;
            END_IF;
        END_IF;

    3: (* East-West Yellow *)
        EastWestYellow := TRUE;
        NorthSouthRed := TRUE;
        Timer(IN := TRUE, PT := T#2s); (* Yellow light duration *)
        IF Timer.Q THEN
            Timer(IN := FALSE);
            LightState := 0;
        END_IF;

END_CASE;

END_FUNCTION_BLOCK

(* ---- M128.st ---- *)
FUNCTION_BLOCK TRAFFIC_CTRL

VAR_INPUT
    PedestrianButton1 : BOOL;
    PedestrianButton2 : BOOL;
END_VAR

VAR_OUTPUT
    NorthSouthRed : BOOL;
    NorthSouthYellow : BOOL;
    NorthSouthGreen : BOOL;
    EastWestRed : BOOL;
    EastWestYellow : BOOL;
    EastWestGreen : BOOL;
    PedestrianLight1 : BOOL;
    PedestrianLight2 : BOOL;
END_VAR

VAR
    LightState : INT := 0; (* 0: North-South Green, 1: North-South Yellow, 2: East-West Green, 3: East-West Yellow *)
    PedestrianRequest1 : BOOL := FALSE;
    PedestrianRequest2 : BOOL := FALSE;
    PedestrianCrossing : BOOL := FALSE;
    Timer : TON;
END_VAR

(* Check for pedestrian requests *)
IF PedestrianButton1 THEN
    PedestrianRequest1 := TRUE;
END_IF;

IF PedestrianButton2 THEN
    PedestrianRequest2 := TRUE;
END_IF;

(* Traffic light state machine *)
CASE LightState OF
    0: (* North-South Green *)
        NorthSouthGreen := TRUE;
        EastWestRed := TRUE;
        IF PedestrianRequest1 OR PedestrianRequest2 THEN
            Timer(IN := TRUE, PT := T#2s); (* Pedestrian crossing grace period *)
            IF Timer.Q THEN
                Timer(IN := FALSE);
                LightState := 1;
            END_IF;
        END_IF;

    1: (* North-South Yellow *)
        NorthSouthYellow := TRUE;
        EastWestRed := TRUE;
        Timer(IN := TRUE, PT := T#2s); (* Yellow light duration *)
        IF Timer.Q THEN
            Timer(IN := FALSE);
            LightState := 2;
        END_IF;

    2: (* East-West Green *)
        EastWestGreen := TRUE;
        NorthSouthRed := TRUE;
        IF PedestrianRequest1 THEN
            PedestrianLight1 := TRUE;
            PedestrianCrossing := TRUE;
        END_IF;
        IF PedestrianRequest2 THEN
            PedestrianLight2 := TRUE;
            PedestrianCrossing := TRUE;
        END_IF;
        IF PedestrianCrossing THEN
            Timer(IN := TRUE, PT := T#2s); (* Pedestrian crossing period *)
            IF Timer.Q THEN
                Timer(IN := FALSE);
                PedestrianRequest1 := FALSE;
                PedestrianRequest2 := FALSE;
                PedestrianLight1 := FALSE;
                PedestrianLight2 := FALSE;
                PedestrianCrossing := FALSE;
                LightState := 3;
            END_IF;
        END_IF;

    3: (* East-West Yellow *)
        EastWestYellow := FALSE; (* MUTATED: BOOL_CONST_REPLACE *)
        NorthSouthRed := TRUE;
        Timer(IN := TRUE, PT := T#2s); (* Yellow light duration *)
        IF Timer.Q THEN
            Timer(IN := FALSE);
            LightState := 0;
        END_IF;

END_CASE;

END_FUNCTION_BLOCK

(* ---- M129.st ---- *)
FUNCTION_BLOCK TRAFFIC_CTRL

VAR_INPUT
    PedestrianButton1 : BOOL;
    PedestrianButton2 : BOOL;
END_VAR

VAR_OUTPUT
    NorthSouthRed : BOOL;
    NorthSouthYellow : BOOL;
    NorthSouthGreen : BOOL;
    EastWestRed : BOOL;
    EastWestYellow : BOOL;
    EastWestGreen : BOOL;
    PedestrianLight1 : BOOL;
    PedestrianLight2 : BOOL;
END_VAR

VAR
    LightState : INT := 0; (* 0: North-South Green, 1: North-South Yellow, 2: East-West Green, 3: East-West Yellow *)
    PedestrianRequest1 : BOOL := FALSE;
    PedestrianRequest2 : BOOL := FALSE;
    PedestrianCrossing : BOOL := FALSE;
    Timer : TON;
END_VAR

(* Check for pedestrian requests *)
IF PedestrianButton1 THEN
    PedestrianRequest1 := TRUE;
END_IF;

IF PedestrianButton2 THEN
    PedestrianRequest2 := TRUE;
END_IF;

(* Traffic light state machine *)
CASE LightState OF
    0: (* North-South Green *)
        NorthSouthGreen := TRUE;
        EastWestRed := TRUE;
        IF PedestrianRequest1 OR PedestrianRequest2 THEN
            Timer(IN := TRUE, PT := T#2s); (* Pedestrian crossing grace period *)
            IF Timer.Q THEN
                Timer(IN := FALSE);
                LightState := 1;
            END_IF;
        END_IF;

    1: (* North-South Yellow *)
        NorthSouthYellow := TRUE;
        EastWestRed := TRUE;
        Timer(IN := TRUE, PT := T#2s); (* Yellow light duration *)
        IF Timer.Q THEN
            Timer(IN := FALSE);
            LightState := 2;
        END_IF;

    2: (* East-West Green *)
        EastWestGreen := TRUE;
        NorthSouthRed := TRUE;
        IF PedestrianRequest1 THEN
            PedestrianLight1 := TRUE;
            PedestrianCrossing := TRUE;
        END_IF;
        IF PedestrianRequest2 THEN
            PedestrianLight2 := TRUE;
            PedestrianCrossing := TRUE;
        END_IF;
        IF PedestrianCrossing THEN
            Timer(IN := TRUE, PT := T#2s); (* Pedestrian crossing period *)
            IF Timer.Q THEN
                Timer(IN := FALSE);
                PedestrianRequest1 := FALSE;
                PedestrianRequest2 := FALSE;
                PedestrianLight1 := FALSE;
                PedestrianLight2 := FALSE;
                PedestrianCrossing := FALSE;
                LightState := 3;
            END_IF;
        END_IF;

    3: (* East-West Yellow *)
        EastWestYellow := TRUE;
        NorthSouthRed := FALSE; (* MUTATED: BOOL_CONST_REPLACE *)
        Timer(IN := TRUE, PT := T#2s); (* Yellow light duration *)
        IF Timer.Q THEN
            Timer(IN := FALSE);
            LightState := 0;
        END_IF;

END_CASE;

END_FUNCTION_BLOCK

(* ---- M130.st ---- *)
FUNCTION_BLOCK TRAFFIC_CTRL

VAR_INPUT
    PedestrianButton1 : BOOL;
    PedestrianButton2 : BOOL;
END_VAR

VAR_OUTPUT
    NorthSouthRed : BOOL;
    NorthSouthYellow : BOOL;
    NorthSouthGreen : BOOL;
    EastWestRed : BOOL;
    EastWestYellow : BOOL;
    EastWestGreen : BOOL;
    PedestrianLight1 : BOOL;
    PedestrianLight2 : BOOL;
END_VAR

VAR
    LightState : INT := 0; (* 0: North-South Green, 1: North-South Yellow, 2: East-West Green, 3: East-West Yellow *)
    PedestrianRequest1 : BOOL := FALSE;
    PedestrianRequest2 : BOOL := FALSE;
    PedestrianCrossing : BOOL := FALSE;
    Timer : TON;
END_VAR

(* Check for pedestrian requests *)
IF PedestrianButton1 THEN
    PedestrianRequest1 := TRUE;
END_IF;

IF PedestrianButton2 THEN
    PedestrianRequest2 := TRUE;
END_IF;

(* Traffic light state machine *)
CASE LightState OF
    0: (* North-South Green *)
        NorthSouthGreen := TRUE;
        EastWestRed := TRUE;
        IF PedestrianRequest1 OR PedestrianRequest2 THEN
            Timer(IN := TRUE, PT := T#2s); (* Pedestrian crossing grace period *)
            IF Timer.Q THEN
                Timer(IN := FALSE);
                LightState := 1;
            END_IF;
        END_IF;

    1: (* North-South Yellow *)
        NorthSouthYellow := TRUE;
        EastWestRed := TRUE;
        Timer(IN := TRUE, PT := T#2s); (* Yellow light duration *)
        IF Timer.Q THEN
            Timer(IN := FALSE);
            LightState := 2;
        END_IF;

    2: (* East-West Green *)
        EastWestGreen := TRUE;
        NorthSouthRed := TRUE;
        IF PedestrianRequest1 THEN
            PedestrianLight1 := TRUE;
            PedestrianCrossing := TRUE;
        END_IF;
        IF PedestrianRequest2 THEN
            PedestrianLight2 := TRUE;
            PedestrianCrossing := TRUE;
        END_IF;
        IF PedestrianCrossing THEN
            Timer(IN := TRUE, PT := T#2s); (* Pedestrian crossing period *)
            IF Timer.Q THEN
                Timer(IN := FALSE);
                PedestrianRequest1 := FALSE;
                PedestrianRequest2 := FALSE;
                PedestrianLight1 := FALSE;
                PedestrianLight2 := FALSE;
                PedestrianCrossing := FALSE;
                LightState := 3;
            END_IF;
        END_IF;

    3: (* East-West Yellow *)
        EastWestYellow := TRUE;
        NorthSouthRed := TRUE;
        Timer(IN := FALSE, PT := T#2s); (* Yellow light duration *) (* MUTATED: BOOL_CONST_REPLACE *)
        IF Timer.Q THEN
            Timer(IN := FALSE);
            LightState := 0;
        END_IF;

END_CASE;

END_FUNCTION_BLOCK

(* ---- M131.st ---- *)
FUNCTION_BLOCK TRAFFIC_CTRL

VAR_INPUT
    PedestrianButton1 : BOOL;
    PedestrianButton2 : BOOL;
END_VAR

VAR_OUTPUT
    NorthSouthRed : BOOL;
    NorthSouthYellow : BOOL;
    NorthSouthGreen : BOOL;
    EastWestRed : BOOL;
    EastWestYellow : BOOL;
    EastWestGreen : BOOL;
    PedestrianLight1 : BOOL;
    PedestrianLight2 : BOOL;
END_VAR

VAR
    LightState : INT := 0; (* 0: North-South Green, 1: North-South Yellow, 2: East-West Green, 3: East-West Yellow *)
    PedestrianRequest1 : BOOL := FALSE;
    PedestrianRequest2 : BOOL := FALSE;
    PedestrianCrossing : BOOL := FALSE;
    Timer : TON;
END_VAR

(* Check for pedestrian requests *)
IF PedestrianButton1 THEN
    PedestrianRequest1 := TRUE;
END_IF;

IF PedestrianButton2 THEN
    PedestrianRequest2 := TRUE;
END_IF;

(* Traffic light state machine *)
CASE LightState OF
    0: (* North-South Green *)
        NorthSouthGreen := TRUE;
        EastWestRed := TRUE;
        IF PedestrianRequest1 OR PedestrianRequest2 THEN
            Timer(IN := TRUE, PT := T#2s); (* Pedestrian crossing grace period *)
            IF Timer.Q THEN
                Timer(IN := FALSE);
                LightState := 1;
            END_IF;
        END_IF;

    1: (* North-South Yellow *)
        NorthSouthYellow := TRUE;
        EastWestRed := TRUE;
        Timer(IN := TRUE, PT := T#2s); (* Yellow light duration *)
        IF Timer.Q THEN
            Timer(IN := FALSE);
            LightState := 2;
        END_IF;

    2: (* East-West Green *)
        EastWestGreen := TRUE;
        NorthSouthRed := TRUE;
        IF PedestrianRequest1 THEN
            PedestrianLight1 := TRUE;
            PedestrianCrossing := TRUE;
        END_IF;
        IF PedestrianRequest2 THEN
            PedestrianLight2 := TRUE;
            PedestrianCrossing := TRUE;
        END_IF;
        IF PedestrianCrossing THEN
            Timer(IN := TRUE, PT := T#2s); (* Pedestrian crossing period *)
            IF Timer.Q THEN
                Timer(IN := FALSE);
                PedestrianRequest1 := FALSE;
                PedestrianRequest2 := FALSE;
                PedestrianLight1 := FALSE;
                PedestrianLight2 := FALSE;
                PedestrianCrossing := FALSE;
                LightState := 3;
            END_IF;
        END_IF;

    3: (* East-West Yellow *)
        EastWestYellow := TRUE;
        NorthSouthRed := TRUE;
        Timer(IN := TRUE, PT := T#2s); (* Yellow light duration *)
        IF Timer.Q THEN
            Timer(IN := TRUE); (* MUTATED: BOOL_CONST_REPLACE *)
            LightState := 0;
        END_IF;

END_CASE;

END_FUNCTION_BLOCK

(* ---- M132.st ---- *)
FUNCTION_BLOCK TRAFFIC_CTRL

VAR_INPUT
    PedestrianButton1 : BOOL;
    PedestrianButton2 : BOOL;
END_VAR

VAR_OUTPUT
    NorthSouthRed : BOOL;
    NorthSouthYellow : BOOL;
    NorthSouthGreen : BOOL;
    EastWestRed : BOOL;
    EastWestYellow : BOOL;
    EastWestGreen : BOOL;
    PedestrianLight1 : BOOL;
    PedestrianLight2 : BOOL;
END_VAR

VAR
    LightState : INT := 0; (* 0: North-South Green, 1: North-South Yellow, 2: East-West Green, 3: East-West Yellow *)
    PedestrianRequest1 : BOOL := FALSE;
    PedestrianRequest2 : BOOL := FALSE;
    PedestrianCrossing : BOOL := FALSE;
    Timer : TON;
END_VAR

(* Check for pedestrian requests *)
IF PedestrianButton1 THEN
    PedestrianRequest1 := TRUE;
END_IF;

IF PedestrianButton2 THEN
    PedestrianRequest2 := TRUE;
END_IF;

(* Traffic light state machine *)
CASE LightState OF
    1: (* North-South Green *) (* MUTATED: CONST_VALUE_REPLACE *)
        NorthSouthGreen := TRUE;
        EastWestRed := TRUE;
        IF PedestrianRequest1 OR PedestrianRequest2 THEN
            Timer(IN := TRUE, PT := T#2s); (* Pedestrian crossing grace period *)
            IF Timer.Q THEN
                Timer(IN := FALSE);
                LightState := 1;
            END_IF;
        END_IF;

    1: (* North-South Yellow *)
        NorthSouthYellow := TRUE;
        EastWestRed := TRUE;
        Timer(IN := TRUE, PT := T#2s); (* Yellow light duration *)
        IF Timer.Q THEN
            Timer(IN := FALSE);
            LightState := 2;
        END_IF;

    2: (* East-West Green *)
        EastWestGreen := TRUE;
        NorthSouthRed := TRUE;
        IF PedestrianRequest1 THEN
            PedestrianLight1 := TRUE;
            PedestrianCrossing := TRUE;
        END_IF;
        IF PedestrianRequest2 THEN
            PedestrianLight2 := TRUE;
            PedestrianCrossing := TRUE;
        END_IF;
        IF PedestrianCrossing THEN
            Timer(IN := TRUE, PT := T#2s); (* Pedestrian crossing period *)
            IF Timer.Q THEN
                Timer(IN := FALSE);
                PedestrianRequest1 := FALSE;
                PedestrianRequest2 := FALSE;
                PedestrianLight1 := FALSE;
                PedestrianLight2 := FALSE;
                PedestrianCrossing := FALSE;
                LightState := 3;
            END_IF;
        END_IF;

    3: (* East-West Yellow *)
        EastWestYellow := TRUE;
        NorthSouthRed := TRUE;
        Timer(IN := TRUE, PT := T#2s); (* Yellow light duration *)
        IF Timer.Q THEN
            Timer(IN := FALSE);
            LightState := 0;
        END_IF;

END_CASE;

END_FUNCTION_BLOCK
